(* IEC 61131-3 sources: plc-st-coding-agent/progress/evidence/f14_v14_remaining_20261113/jobs/codex_minimax-m27 (part 5) *)

(* ---- self-hard-03.raw_candidate_01.st ---- *)
(* ENGINEERING_CONTRACT
 * FIFO Queue with 8-slot compact array
 * [PUB001-PUB010] Core ops: popEn rising→remove first if count>0; pushEn rising→add pushItem if count<8
 *   Same-scan priority: pop executes BEFORE push; full→pop+push (net 0), empty→push-only (net +1)
 * [PUB011] Retention: count and fifo[1..8] state retained in VAR between scans
 * [PUB012] No AT located declarations
 * [PUB013-PUB015] Rising edge: each button triggers once per press; initial history=FALSE
 * [PUB016-PUB019] Same-scan semantics: full queue drains one slot then accepts push; empty queue accepts push only
 * [PUB020-PUB025] Array bounds: fifo[1..8], compact at end of scan: fifo[1..count] is logical queue FIFO order
 *   head=fifo[1] when non-empty, else 0; fifo[count+1..8] unspecified/unconstrained
 * [PUB026-PUB030] count∈[0,8], full↔count=8, empty↔count=0; success of push/pop updates count
 *)

(* CONTRACT_RULES [] *)

FUNCTION_BLOCK FB
VAR_INPUT
    pushEn    : BOOL;
    pushItem  : INT;
    popEn     : BOOL;
END_VAR
VAR_IN_OUT
    fifo      : ARRAY[1..8] OF INT;
END_VAR
VAR_OUTPUT
    count     : INT;
    full      : BOOL;
    empty     : BOOL;
    head      : INT;
END_VAR
VAR
    prev_pushEn : BOOL := FALSE;
    prev_popEn  : BOOL := FALSE;
    tmp_pushRising : BOOL;
    tmp_popRising  : BOOL;
    tmp_i       : INT;
END_VAR

    // Rising edge detection
    tmp_popRising  := popEn AND NOT prev_popEn;
    tmp_pushRising := pushEn AND NOT prev_pushEn;
    prev_popEn  := popEn;
    prev_pushEn := pushEn;

    // Execute in required order: pop first, then push
    // POP: non-empty queue only
    IF tmp_popRising AND count > 0 THEN
        FOR tmp_i := 1 TO count - 1 DO
            fifo[tmp_i] := fifo[tmp_i + 1];
        END_FOR;
        count := count - 1;
    END_IF;

    // PUSH: non-full queue only
    IF tmp_pushRising AND count < 8 THEN
        count := count + 1;
        fifo[count] := pushItem;
    END_IF;

    // Outputs
    full  := (count = 8);
    empty := (count = 0);
    IF empty THEN
        head := 0;
    ELSE
        head := fifo[1];
    END_IF;

END_FUNCTION_BLOCK

(* ---- self-hard-04.candidate_01.st ---- *)
(*
ENGINEERING_CONTRACT
==================
State retention & activation:
- leadPump: latches until demand=0 clears it; reset_input=demand<=0 PUB004
- lagPump: latches until demand<2 clears it; hold on same-scan no-rise PUB005
- runningCount: combinational, equals clipped demand every scan PUB001
Initialization:
- First positive demand after demand=0 selects shortest-run pump as leadPump (PUB010)
- First positive demand sets lagPump if demand>=2 (PUB011)
Rotation behavior:
- rotated=TRUE + main.runHours - MIN(runHours) > 50 → switch to shortest (PUB012)
- rotated=FALSE → never switch, even if hysteresis gap exists (PUB012)
- rotated is level-triggered, evaluated every scan with current main hours (PUB012)
Backup selection moments:
- Initial selection | leadPump change | runningCount increase → recompute lagPump (PUB026)
- Otherwise retain previous lagPump (PUB028)
Direction conflict: N/A (no opposite movements in this pump-selection task)
Units: runHours in LINT hours, 50-hour hysteresis threshold (PUB012)
*)
(* CONTRACT_RULES [] *)

FUNCTION_BLOCK FB
VAR_INPUT
    demand     : INT;
    runHours   : ARRAY[1..5] OF LINT;
    rotated    : BOOL;
END_VAR
VAR_OUTPUT
    leadPump   : INT := 0;
    lagPump    : INT := 0;
    runningCount : INT := 0;
END_VAR
VAR
    prevLeadPump    : INT := 0;
    prevLagPump     : INT := 0;
    prevRunningCount : INT := 0;
    prevClippedDemand : INT := 0;
    wasDemandZero   : BOOL := TRUE;
END_VAR

VAR
    clippedDemand : INT;
    tmp_i         : INT;
    tmp_minHours  : LINT;
    tmp_minPump   : INT;
    tmp_secondMinHours : LINT;
    tmp_secondMinPump  : INT;
    tmp_mainHoursDiff  : LINT;
END_VAR

    // PUB001: Clip demand to 0..5
    IF demand < 0 THEN
        clippedDemand := 0;
    ELSIF demand > 5 THEN
        clippedDemand := 5;
    ELSE
        clippedDemand := demand;
    END_IF;

    runningCount := clippedDemand;

    // Clear all outputs when demand <= 0
    IF clippedDemand = 0 THEN
        leadPump := 0;
        lagPump  := 0;
        prevLeadPump    := 0;
        prevLagPump     := 0;
        prevRunningCount := 0;
        prevClippedDemand := 0;
        wasDemandZero   := TRUE;
    ELSE
        // Find pump with minimum run hours (for hysteresis check and selection)
        tmp_minHours := runHours[1];
        tmp_minPump  := 1;
        FOR tmp_i := 2 TO 5 DO
            IF runHours[tmp_i] < tmp_minHours THEN
                tmp_minHours := runHours[tmp_i];
                tmp_minPump  := tmp_i;
            ELSIF runHours[tmp_i] = tmp_minHours AND tmp_i < tmp_minPump THEN
                tmp_minPump  := tmp_i;
            END_IF;
        END_FOR;

        // Determine if this is initial selection (first positive demand after zero)
        IF wasDemandZero THEN
            // Initial selection: pick shortest-run pump as main
            leadPump   := tmp_minPump;
            lagPump    := 0;
            wasDemandZero := FALSE;
        ELSE
            // Not initial selection: check for rotation request
            IF rotated AND prevLeadPump <> 0 THEN
                // Compute main pump's hours difference from minimum
                tmp_mainHoursDiff := runHours[prevLeadPump] - tmp_minHours;
                IF tmp_mainHoursDiff > 50 THEN
                    // Hysteresis satisfied: switch to shortest-run pump
                    leadPump := tmp_minPump;
                ELSE
                    // Keep current main pump
                    leadPump := prevLeadPump;
                END_IF;
            ELSE
                // No rotation request or no previous main: keep current main
                leadPump := prevLeadPump;
            END_IF;
        END_IF;

        // Backup pump selection (PUB026, PUB028)
        IF clippedDemand >= 2 THEN
            // Need backup pump
            // Recompute lagPump only on: initial, leadPump change, runningCount increase
            IF wasDemandZero OR leadPump <> prevLeadPump OR clippedDemand > prevClippedDemand THEN
                // Find second-minimum pump (excluding leadPump)
                tmp_secondMinHours := 16#7FFFFFFFFFFFFFFF; // Large LINT value
                tmp_secondMinPump  := 0;
                FOR tmp_i := 1 TO 5 DO
                    IF tmp_i = leadPump THEN
                        // Skip main pump
                    ELSE
                        IF runHours[tmp_i] < tmp_secondMinHours THEN
                            tmp_secondMinHours := runHours[tmp_i];
                            tmp_secondMinPump  := tmp_i;
                        ELSIF runHours[tmp_i] = tmp_secondMinHours AND tmp_i < tmp_secondMinPump THEN
                            tmp_secondMinPump  := tmp_i;
                        END_IF;
                    END_IF;
                END_FOR;
                lagPump := tmp_secondMinPump;
            ELSE
                // Retain previous backup pump
                lagPump := prevLagPump;
            END_IF;
        ELSE
            // Demand < 2: no backup pump
            lagPump := 0;
        END_IF;
    END_IF;

    // Update previous state for next scan
    prevLeadPump     := leadPump;
    prevLagPump      := lagPump;
    prevRunningCount := runningCount;
    prevClippedDemand := clippedDemand;

END_FUNCTION_BLOCK

(* ---- self-hard-04.candidate_03.st ---- *)
(*
ENGINEERING_CONTRACT
==================
State retention & activation:
- leadPump: latches until demand=0 clears it; reset_input=demand<=0 PUB004
- lagPump: latches until demand<2 clears it; hold on same-scan no-rise PUB005
- runningCount: combinational, equals clipped demand every scan PUB001
Initialization:
- First positive demand after demand=0 selects shortest-run pump as leadPump (PUB010)
- First positive demand sets lagPump if demand>=2 (PUB011)
Rotation behavior:
- rotated=TRUE + main.runHours - MIN(runHours) > 50 → switch to shortest (PUB012)
- rotated=FALSE → never switch, even if hysteresis gap exists (PUB012)
- rotated is level-triggered, evaluated every scan with current main hours (PUB012)
Backup selection moments:
- Initial selection | leadPump change | runningCount increase → recompute lagPump (PUB026)
- Otherwise retain previous lagPump (PUB028)
Direction conflict: N/A (no opposite movements in this pump-selection task)
Units: runHours in LINT hours, 50-hour hysteresis threshold (PUB012)
*)
(* CONTRACT_RULES [] *)

FUNCTION_BLOCK FB
VAR_INPUT
    demand     : INT;
    runHours   : ARRAY[1..5] OF LINT;
    rotated    : BOOL;
END_VAR
VAR_OUTPUT
    leadPump   : INT := 0;
    lagPump    : INT := 0;
    runningCount : INT := 0;
END_VAR
VAR
    prevLeadPump    : INT := 0;
    prevLagPump     : INT := 0;
    prevRunningCount : INT := 0;
    prevClippedDemand : INT := 0;
    wasDemandZero   : BOOL := TRUE;
    clippedDemand : INT;
    tmp_i         : INT;
    tmp_minHours  : LINT;
    tmp_minPump   : INT;
    tmp_secondMinHours : LINT;
    tmp_secondMinPump  : INT;
    tmp_mainHoursDiff  : LINT;
END_VAR

    // PUB001: Clip demand to 0..5
    IF demand < 0 THEN
        clippedDemand := 0;
    ELSIF demand > 5 THEN
        clippedDemand := 5;
    ELSE
        clippedDemand := demand;
    END_IF;

    runningCount := clippedDemand;

    // Clear all outputs when demand <= 0
    IF clippedDemand = 0 THEN
        leadPump := 0;
        lagPump  := 0;
        prevLeadPump    := 0;
        prevLagPump     := 0;
        prevRunningCount := 0;
        prevClippedDemand := 0;
        wasDemandZero   := TRUE;
    ELSE
        // Find pump with minimum run hours (for hysteresis check and selection)
        tmp_minHours := runHours[1];
        tmp_minPump  := 1;
        FOR tmp_i := 2 TO 5 DO
            IF runHours[tmp_i] < tmp_minHours THEN
                tmp_minHours := runHours[tmp_i];
                tmp_minPump  := tmp_i;
            ELSIF runHours[tmp_i] = tmp_minHours AND tmp_i < tmp_minPump THEN
                tmp_minPump  := tmp_i;
            END_IF;
        END_FOR;

        // Determine if this is initial selection (first positive demand after zero)
        IF wasDemandZero THEN
            // Initial selection: pick shortest-run pump as main
            leadPump   := tmp_minPump;
            lagPump    := 0;
            wasDemandZero := FALSE;
        ELSE
            // Not initial selection: check for rotation request
            IF rotated AND prevLeadPump <> 0 THEN
                // Compute main pump's hours difference from minimum
                tmp_mainHoursDiff := runHours[prevLeadPump] - tmp_minHours;
                IF tmp_mainHoursDiff > 50 THEN
                    // Hysteresis satisfied: switch to shortest-run pump
                    leadPump := tmp_minPump;
                ELSE
                    // Keep current main pump
                    leadPump := prevLeadPump;
                END_IF;
            ELSE
                // No rotation request or no previous main: keep current main
                leadPump := prevLeadPump;
            END_IF;
        END_IF;

        // Backup pump selection (PUB026, PUB028)
        IF clippedDemand >= 2 THEN
            // Need backup pump
            // Recompute lagPump only on: initial, leadPump change, runningCount increase
            IF wasDemandZero OR leadPump <> prevLeadPump OR clippedDemand > prevClippedDemand THEN
                // Find second-minimum pump (excluding leadPump)
                tmp_secondMinHours := 16#7FFFFFFFFFFFFFFF; // Large LINT value
                tmp_secondMinPump  := 0;
                FOR tmp_i := 1 TO 5 DO
                    IF tmp_i = leadPump THEN
                        // Skip main pump
                    ELSE
                        IF runHours[tmp_i] < tmp_secondMinHours THEN
                            tmp_secondMinHours := runHours[tmp_i];
                            tmp_secondMinPump  := tmp_i;
                        ELSIF runHours[tmp_i] = tmp_secondMinHours AND tmp_i < tmp_secondMinPump THEN
                            tmp_secondMinPump  := tmp_i;
                        END_IF;
                    END_IF;
                END_FOR;
                lagPump := tmp_secondMinPump;
            ELSE
                // Retain previous backup pump
                lagPump := prevLagPump;
            END_IF;
        ELSE
            // Demand < 2: no backup pump
            lagPump := 0;
        END_IF;
    END_IF;

    // Update previous state for next scan
    prevLeadPump     := leadPump;
    prevLagPump      := lagPump;
    prevRunningCount := runningCount;
    prevClippedDemand := clippedDemand;

END_FUNCTION_BLOCK

(* ---- self-hard-04.patch_base_02.st ---- *)
(*
ENGINEERING_CONTRACT
==================
State retention & activation:
- leadPump: latches until demand=0 clears it; reset_input=demand<=0 PUB004
- lagPump: latches until demand<2 clears it; hold on same-scan no-rise PUB005
- runningCount: combinational, equals clipped demand every scan PUB001
Initialization:
- First positive demand after demand=0 selects shortest-run pump as leadPump (PUB010)
- First positive demand sets lagPump if demand>=2 (PUB011)
Rotation behavior:
- rotated=TRUE + main.runHours - MIN(runHours) > 50 → switch to shortest (PUB012)
- rotated=FALSE → never switch, even if hysteresis gap exists (PUB012)
- rotated is level-triggered, evaluated every scan with current main hours (PUB012)
Backup selection moments:
- Initial selection | leadPump change | runningCount increase → recompute lagPump (PUB026)
- Otherwise retain previous lagPump (PUB028)
Direction conflict: N/A (no opposite movements in this pump-selection task)
Units: runHours in LINT hours, 50-hour hysteresis threshold (PUB012)
*)
(* CONTRACT_RULES [] *)

FUNCTION_BLOCK FB
VAR_INPUT
    demand     : INT;
    runHours   : ARRAY[1..5] OF LINT;
    rotated    : BOOL;
END_VAR
VAR_OUTPUT
    leadPump   : INT := 0;
    lagPump    : INT := 0;
    runningCount : INT := 0;
END_VAR
VAR
    prevLeadPump    : INT := 0;
    prevLagPump     : INT := 0;
    prevRunningCount : INT := 0;
    prevClippedDemand : INT := 0;
    wasDemandZero   : BOOL := TRUE;
END_VAR

VAR
    clippedDemand : INT;
    tmp_i         : INT;
    tmp_minHours  : LINT;
    tmp_minPump   : INT;
    tmp_secondMinHours : LINT;
    tmp_secondMinPump  : INT;
    tmp_mainHoursDiff  : LINT;
END_VAR

    // PUB001: Clip demand to 0..5
    IF demand < 0 THEN
        clippedDemand := 0;
    ELSIF demand > 5 THEN
        clippedDemand := 5;
    ELSE
        clippedDemand := demand;
    END_IF;

    runningCount := clippedDemand;

    // Clear all outputs when demand <= 0
    IF clippedDemand = 0 THEN
        leadPump := 0;
        lagPump  := 0;
        prevLeadPump    := 0;
        prevLagPump     := 0;
        prevRunningCount := 0;
        prevClippedDemand := 0;
        wasDemandZero   := TRUE;
    ELSE
        // Find pump with minimum run hours (for hysteresis check and selection)
        tmp_minHours := runHours[1];
        tmp_minPump  := 1;
        FOR tmp_i := 2 TO 5 DO
            IF runHours[tmp_i] < tmp_minHours THEN
                tmp_minHours := runHours[tmp_i];
                tmp_minPump  := tmp_i;
            ELSIF runHours[tmp_i] = tmp_minHours AND tmp_i < tmp_minPump THEN
                tmp_minPump  := tmp_i;
            END_IF;
        END_FOR;

        // Determine if this is initial selection (first positive demand after zero)
        IF wasDemandZero THEN
            // Initial selection: pick shortest-run pump as main
            leadPump   := tmp_minPump;
            lagPump    := 0;
            wasDemandZero := FALSE;
        ELSE
            // Not initial selection: check for rotation request
            IF rotated AND prevLeadPump <> 0 THEN
                // Compute main pump's hours difference from minimum
                tmp_mainHoursDiff := runHours[prevLeadPump] - tmp_minHours;
                IF tmp_mainHoursDiff > 50 THEN
                    // Hysteresis satisfied: switch to shortest-run pump
                    leadPump := tmp_minPump;
                ELSE
                    // Keep current main pump
                    leadPump := prevLeadPump;
                END_IF;
            ELSE
                // No rotation request or no previous main: keep current main
                leadPump := prevLeadPump;
            END_IF;
        END_IF;

        // Backup pump selection (PUB026, PUB028)
        IF clippedDemand >= 2 THEN
            // Need backup pump
            // Recompute lagPump only on: initial, leadPump change, runningCount increase
            IF wasDemandZero OR leadPump <> prevLeadPump OR clippedDemand > prevClippedDemand THEN
                // Find second-minimum pump (excluding leadPump)
                tmp_secondMinHours := 16#7FFFFFFFFFFFFFFF; // Large LINT value
                tmp_secondMinPump  := 0;
                FOR tmp_i := 1 TO 5 DO
                    IF tmp_i = leadPump THEN
                        // Skip main pump
                    ELSE
                        IF runHours[tmp_i] < tmp_secondMinHours THEN
                            tmp_secondMinHours := runHours[tmp_i];
                            tmp_secondMinPump  := tmp_i;
                        ELSIF runHours[tmp_i] = tmp_secondMinHours AND tmp_i < tmp_secondMinPump THEN
                            tmp_secondMinPump  := tmp_i;
                        END_IF;
                    END_IF;
                END_FOR;
                lagPump := tmp_secondMinPump;
            ELSE
                // Retain previous backup pump
                lagPump := prevLagPump;
            END_IF;
        ELSE
            // Demand < 2: no backup pump
            lagPump := 0;
        END_IF;
    END_IF;

    // Update previous state for next scan
    prevLeadPump     := leadPump;
    prevLagPump      := lagPump;
    prevRunningCount := runningCount;
    prevClippedDemand := clippedDemand;

END_FUNCTION_BLOCK

(* ---- self-hard-04.patch_base_03.st ---- *)
(*
ENGINEERING_CONTRACT
==================
State retention & activation:
- leadPump: latches until demand=0 clears it; reset_input=demand<=0 PUB004
- lagPump: latches until demand<2 clears it; hold on same-scan no-rise PUB005
- runningCount: combinational, equals clipped demand every scan PUB001
Initialization:
- First positive demand after demand=0 selects shortest-run pump as leadPump (PUB010)
- First positive demand sets lagPump if demand>=2 (PUB011)
Rotation behavior:
- rotated=TRUE + main.runHours - MIN(runHours) > 50 → switch to shortest (PUB012)
- rotated=FALSE → never switch, even if hysteresis gap exists (PUB012)
- rotated is level-triggered, evaluated every scan with current main hours (PUB012)
Backup selection moments:
- Initial selection | leadPump change | runningCount increase → recompute lagPump (PUB026)
- Otherwise retain previous lagPump (PUB028)
Direction conflict: N/A (no opposite movements in this pump-selection task)
Units: runHours in LINT hours, 50-hour hysteresis threshold (PUB012)
*)
(* CONTRACT_RULES [] *)

FUNCTION_BLOCK FB
VAR_INPUT
    demand     : INT;
    runHours   : ARRAY[1..5] OF LINT;
    rotated    : BOOL;
END_VAR
VAR_OUTPUT
    leadPump   : INT := 0;
    lagPump    : INT := 0;
    runningCount : INT := 0;
END_VAR
VAR
    prevLeadPump    : INT := 0;
    prevLagPump     : INT := 0;
    prevRunningCount : INT := 0;
    prevClippedDemand : INT := 0;
    wasDemandZero   : BOOL := TRUE;
END_VAR

VAR
    clippedDemand : INT;
    tmp_i         : INT;
    tmp_minHours  : LINT;
    tmp_minPump   : INT;
    tmp_secondMinHours : LINT;
    tmp_secondMinPump  : INT;
    tmp_mainHoursDiff  : LINT;
END_VAR

    // PUB001: Clip demand to 0..5
    IF demand < 0 THEN
        clippedDemand := 0;
    ELSIF demand > 5 THEN
        clippedDemand := 5;
    ELSE
        clippedDemand := demand;
    END_IF;

    runningCount := clippedDemand;

    // Clear all outputs when demand <= 0
    IF clippedDemand = 0 THEN
        leadPump := 0;
        lagPump  := 0;
        prevLeadPump    := 0;
        prevLagPump     := 0;
        prevRunningCount := 0;
        prevClippedDemand := 0;
        wasDemandZero   := TRUE;
    ELSE
        // Find pump with minimum run hours (for hysteresis check and selection)
        tmp_minHours := runHours[1];
        tmp_minPump  := 1;
        FOR tmp_i := 2 TO 5 DO
            IF runHours[tmp_i] < tmp_minHours THEN
                tmp_minHours := runHours[tmp_i];
                tmp_minPump  := tmp_i;
            ELSIF runHours[tmp_i] = tmp_minHours AND tmp_i < tmp_minPump THEN
                tmp_minPump  := tmp_i;
            END_IF;
        END_FOR;

        // Determine if this is initial selection (first positive demand after zero)
        IF wasDemandZero THEN
            // Initial selection: pick shortest-run pump as main
            leadPump   := tmp_minPump;
            lagPump    := 0;
            wasDemandZero := FALSE;
        ELSE
            // Not initial selection: check for rotation request
            IF rotated AND prevLeadPump <> 0 THEN
                // Compute main pump's hours difference from minimum
                tmp_mainHoursDiff := runHours[prevLeadPump] - tmp_minHours;
                IF tmp_mainHoursDiff > 50 THEN
                    // Hysteresis satisfied: switch to shortest-run pump
                    leadPump := tmp_minPump;
                ELSE
                    // Keep current main pump
                    leadPump := prevLeadPump;
                END_IF;
            ELSE
                // No rotation request or no previous main: keep current main
                leadPump := prevLeadPump;
            END_IF;
        END_IF;

        // Backup pump selection (PUB026, PUB028)
        IF clippedDemand >= 2 THEN
            // Need backup pump
            // Recompute lagPump only on: initial, leadPump change, runningCount increase
            IF wasDemandZero OR leadPump <> prevLeadPump OR clippedDemand > prevClippedDemand THEN
                // Find second-minimum pump (excluding leadPump)
                tmp_secondMinHours := 16#7FFFFFFFFFFFFFFF; // Large LINT value
                tmp_secondMinPump  := 0;
                FOR tmp_i := 1 TO 5 DO
                    IF tmp_i = leadPump THEN
                        // Skip main pump
                    ELSE
                        IF runHours[tmp_i] < tmp_secondMinHours THEN
                            tmp_secondMinHours := runHours[tmp_i];
                            tmp_secondMinPump  := tmp_i;
                        ELSIF runHours[tmp_i] = tmp_secondMinHours AND tmp_i < tmp_secondMinPump THEN
                            tmp_secondMinPump  := tmp_i;
                        END_IF;
                    END_IF;
                END_FOR;
                lagPump := tmp_secondMinPump;
            ELSE
                // Retain previous backup pump
                lagPump := prevLagPump;
            END_IF;
        ELSE
            // Demand < 2: no backup pump
            lagPump := 0;
        END_IF;
    END_IF;

    // Update previous state for next scan
    prevLeadPump     := leadPump;
    prevLagPump      := lagPump;
    prevRunningCount := runningCount;
    prevClippedDemand := clippedDemand;

END_FUNCTION_BLOCK

(* ---- self-hard-04.patch_base_04.st ---- *)
(*
ENGINEERING_CONTRACT
==================
State retention & activation:
- leadPump: latches until demand=0 clears it; reset_input=demand<=0 PUB004
- lagPump: latches until demand<2 clears it; hold on same-scan no-rise PUB005
- runningCount: combinational, equals clipped demand every scan PUB001
Initialization:
- First positive demand after demand=0 selects shortest-run pump as leadPump (PUB010)
- First positive demand sets lagPump if demand>=2 (PUB011)
Rotation behavior:
- rotated=TRUE + main.runHours - MIN(runHours) > 50 → switch to shortest (PUB012)
- rotated=FALSE → never switch, even if hysteresis gap exists (PUB012)
- rotated is level-triggered, evaluated every scan with current main hours (PUB012)
Backup selection moments:
- Initial selection | leadPump change | runningCount increase → recompute lagPump (PUB026)
- Otherwise retain previous lagPump (PUB028)
Direction conflict: N/A (no opposite movements in this pump-selection task)
Units: runHours in LINT hours, 50-hour hysteresis threshold (PUB012)
*)
(* CONTRACT_RULES [] *)

FUNCTION_BLOCK FB
VAR_INPUT
    demand     : INT;
    runHours   : ARRAY[1..5] OF LINT;
    rotated    : BOOL;
END_VAR
VAR_OUTPUT
    leadPump   : INT := 0;
    lagPump    : INT := 0;
    runningCount : INT := 0;
END_VAR
VAR
    prevLeadPump    : INT := 0;
    prevLagPump     : INT := 0;
    prevRunningCount : INT := 0;
    prevClippedDemand : INT := 0;
    wasDemandZero   : BOOL := TRUE;
    clippedDemand : INT;
    tmp_i         : INT;
    tmp_minHours  : LINT;
    tmp_minPump   : INT;
    tmp_secondMinHours : LINT;
    tmp_secondMinPump  : INT;
    tmp_mainHoursDiff  : LINT;
END_VAR

    // PUB001: Clip demand to 0..5
    IF demand < 0 THEN
        clippedDemand := 0;
    ELSIF demand > 5 THEN
        clippedDemand := 5;
    ELSE
        clippedDemand := demand;
    END_IF;

    runningCount := clippedDemand;

    // Clear all outputs when demand <= 0
    IF clippedDemand = 0 THEN
        leadPump := 0;
        lagPump  := 0;
        prevLeadPump    := 0;
        prevLagPump     := 0;
        prevRunningCount := 0;
        prevClippedDemand := 0;
        wasDemandZero   := TRUE;
    ELSE
        // Find pump with minimum run hours (for hysteresis check and selection)
        tmp_minHours := runHours[1];
        tmp_minPump  := 1;
        FOR tmp_i := 2 TO 5 DO
            IF runHours[tmp_i] < tmp_minHours THEN
                tmp_minHours := runHours[tmp_i];
                tmp_minPump  := tmp_i;
            ELSIF runHours[tmp_i] = tmp_minHours AND tmp_i < tmp_minPump THEN
                tmp_minPump  := tmp_i;
            END_IF;
        END_FOR;

        // Determine if this is initial selection (first positive demand after zero)
        IF wasDemandZero THEN
            // Initial selection: pick shortest-run pump as main
            leadPump   := tmp_minPump;
            lagPump    := 0;
            wasDemandZero := FALSE;
        ELSE
            // Not initial selection: check for rotation request
            IF rotated AND prevLeadPump <> 0 THEN
                // Compute main pump's hours difference from minimum
                tmp_mainHoursDiff := runHours[prevLeadPump] - tmp_minHours;
                IF tmp_mainHoursDiff > 50 THEN
                    // Hysteresis satisfied: switch to shortest-run pump
                    leadPump := tmp_minPump;
                ELSE
                    // Keep current main pump
                    leadPump := prevLeadPump;
                END_IF;
            ELSE
                // No rotation request or no previous main: keep current main
                leadPump := prevLeadPump;
            END_IF;
        END_IF;

        // Backup pump selection (PUB026, PUB028)
        IF clippedDemand >= 2 THEN
            // Need backup pump
            // Recompute lagPump only on: initial, leadPump change, runningCount increase
            IF wasDemandZero OR leadPump <> prevLeadPump OR clippedDemand > prevClippedDemand THEN
                // Find second-minimum pump (excluding leadPump)
                tmp_secondMinHours := 16#7FFFFFFFFFFFFFFF; // Large LINT value
                tmp_secondMinPump  := 0;
                FOR tmp_i := 1 TO 5 DO
                    IF tmp_i = leadPump THEN
                        // Skip main pump
                    ELSE
                        IF runHours[tmp_i] < tmp_secondMinHours THEN
                            tmp_secondMinHours := runHours[tmp_i];
                            tmp_secondMinPump  := tmp_i;
                        ELSIF runHours[tmp_i] = tmp_secondMinHours AND tmp_i < tmp_secondMinPump THEN
                            tmp_secondMinPump  := tmp_i;
                        END_IF;
                    END_IF;
                END_FOR;
                lagPump := tmp_secondMinPump;
            ELSE
                // Retain previous backup pump
                lagPump := prevLagPump;
            END_IF;
        ELSE
            // Demand < 2: no backup pump
            lagPump := 0;
        END_IF;
    END_IF;

    // Update previous state for next scan
    prevLeadPump     := leadPump;
    prevLagPump      := lagPump;
    prevRunningCount := runningCount;
    prevClippedDemand := clippedDemand;

END_FUNCTION_BLOCK

(* ---- self-hard-04.raw_candidate_01.st ---- *)
(*
ENGINEERING_CONTRACT
==================
State retention & activation:
- leadPump: latches until demand=0 clears it; reset_input=demand<=0 PUB004
- lagPump: latches until demand<2 clears it; hold on same-scan no-rise PUB005
- runningCount: combinational, equals clipped demand every scan PUB001
Initialization:
- First positive demand after demand=0 selects shortest-run pump as leadPump (PUB010)
- First positive demand sets lagPump if demand>=2 (PUB011)
Rotation behavior:
- rotated=TRUE + main.runHours - MIN(runHours) > 50 → switch to shortest (PUB012)
- rotated=FALSE → never switch, even if hysteresis gap exists (PUB012)
- rotated is level-triggered, evaluated every scan with current main hours (PUB012)
Backup selection moments:
- Initial selection | leadPump change | runningCount increase → recompute lagPump (PUB026)
- Otherwise retain previous lagPump (PUB028)
Direction conflict: N/A (no opposite movements in this pump-selection task)
Units: runHours in LINT hours, 50-hour hysteresis threshold (PUB012)
*)
(* CONTRACT_RULES [] *)

FUNCTION_BLOCK FB
VAR_INPUT
    demand     : INT;
    runHours   : ARRAY[1..5] OF LINT;
    rotated    : BOOL;
END_VAR
VAR_OUTPUT
    leadPump   : INT := 0;
    lagPump    : INT := 0;
    runningCount : INT := 0;
END_VAR
VAR
    prevLeadPump    : INT := 0;
    prevLagPump     : INT := 0;
    prevRunningCount : INT := 0;
    prevClippedDemand : INT := 0;
    wasDemandZero   : BOOL := TRUE;
END_VAR

VAR
    clippedDemand : INT;
    tmp_i         : INT;
    tmp_minHours  : LINT;
    tmp_minPump   : INT;
    tmp_secondMinHours : LINT;
    tmp_secondMinPump  : INT;
    tmp_mainHoursDiff  : LINT;
END_VAR

    // PUB001: Clip demand to 0..5
    IF demand < 0 THEN
        clippedDemand := 0;
    ELSIF demand > 5 THEN
        clippedDemand := 5;
    ELSE
        clippedDemand := demand;
    END_IF;

    runningCount := clippedDemand;

    // Clear all outputs when demand <= 0
    IF clippedDemand = 0 THEN
        leadPump := 0;
        lagPump  := 0;
        prevLeadPump    := 0;
        prevLagPump     := 0;
        prevRunningCount := 0;
        prevClippedDemand := 0;
        wasDemandZero   := TRUE;
    ELSE
        // Find pump with minimum run hours (for hysteresis check and selection)
        tmp_minHours := runHours[1];
        tmp_minPump  := 1;
        FOR tmp_i := 2 TO 5 DO
            IF runHours[tmp_i] < tmp_minHours THEN
                tmp_minHours := runHours[tmp_i];
                tmp_minPump  := tmp_i;
            ELSIF runHours[tmp_i] = tmp_minHours AND tmp_i < tmp_minPump THEN
                tmp_minPump  := tmp_i;
            END_IF;
        END_FOR;

        // Determine if this is initial selection (first positive demand after zero)
        IF wasDemandZero THEN
            // Initial selection: pick shortest-run pump as main
            leadPump   := tmp_minPump;
            lagPump    := 0;
            wasDemandZero := FALSE;
        ELSE
            // Not initial selection: check for rotation request
            IF rotated AND prevLeadPump <> 0 THEN
                // Compute main pump's hours difference from minimum
                tmp_mainHoursDiff := runHours[prevLeadPump] - tmp_minHours;
                IF tmp_mainHoursDiff > 50 THEN
                    // Hysteresis satisfied: switch to shortest-run pump
                    leadPump := tmp_minPump;
                ELSE
                    // Keep current main pump
                    leadPump := prevLeadPump;
                END_IF;
            ELSE
                // No rotation request or no previous main: keep current main
                leadPump := prevLeadPump;
            END_IF;
        END_IF;

        // Backup pump selection (PUB026, PUB028)
        IF clippedDemand >= 2 THEN
            // Need backup pump
            // Recompute lagPump only on: initial, leadPump change, runningCount increase
            IF wasDemandZero OR leadPump <> prevLeadPump OR clippedDemand > prevClippedDemand THEN
                // Find second-minimum pump (excluding leadPump)
                tmp_secondMinHours := 16#7FFFFFFFFFFFFFFF; // Large LINT value
                tmp_secondMinPump  := 0;
                FOR tmp_i := 1 TO 5 DO
                    IF tmp_i = leadPump THEN
                        // Skip main pump
                    ELSE
                        IF runHours[tmp_i] < tmp_secondMinHours THEN
                            tmp_secondMinHours := runHours[tmp_i];
                            tmp_secondMinPump  := tmp_i;
                        ELSIF runHours[tmp_i] = tmp_secondMinHours AND tmp_i < tmp_secondMinPump THEN
                            tmp_secondMinPump  := tmp_i;
                        END_IF;
                    END_IF;
                END_FOR;
                lagPump := tmp_secondMinPump;
            ELSE
                // Retain previous backup pump
                lagPump := prevLagPump;
            END_IF;
        ELSE
            // Demand < 2: no backup pump
            lagPump := 0;
        END_IF;
    END_IF;

    // Update previous state for next scan
    prevLeadPump     := leadPump;
    prevLagPump      := lagPump;
    prevRunningCount := runningCount;
    prevClippedDemand := clippedDemand;

END_FUNCTION_BLOCK

(* ---- self-hard-04.raw_candidate_03.st ---- *)
(*
ENGINEERING_CONTRACT
==================
State retention & activation:
- leadPump: latches until demand=0 clears it; reset_input=demand<=0 PUB004
- lagPump: latches until demand<2 clears it; hold on same-scan no-rise PUB005
- runningCount: combinational, equals clipped demand every scan PUB001
Initialization:
- First positive demand after demand=0 selects shortest-run pump as leadPump (PUB010)
- First positive demand sets lagPump if demand>=2 (PUB011)
Rotation behavior:
- rotated=TRUE + main.runHours - MIN(runHours) > 50 → switch to shortest (PUB012)
- rotated=FALSE → never switch, even if hysteresis gap exists (PUB012)
- rotated is level-triggered, evaluated every scan with current main hours (PUB012)
Backup selection moments:
- Initial selection | leadPump change | runningCount increase → recompute lagPump (PUB026)
- Otherwise retain previous lagPump (PUB028)
Direction conflict: N/A (no opposite movements in this pump-selection task)
Units: runHours in LINT hours, 50-hour hysteresis threshold (PUB012)
*)
(* CONTRACT_RULES [] *)

FUNCTION_BLOCK FB
VAR_INPUT
    demand     : INT;
    runHours   : ARRAY[1..5] OF LINT;
    rotated    : BOOL;
END_VAR
VAR_OUTPUT
    leadPump   : INT := 0;
    lagPump    : INT := 0;
    runningCount : INT := 0;
END_VAR
VAR
    prevLeadPump    : INT := 0;
    prevLagPump     : INT := 0;
    prevRunningCount : INT := 0;
    prevClippedDemand : INT := 0;
    wasDemandZero   : BOOL := TRUE;
    clippedDemand : INT;
    tmp_i         : INT;
    tmp_minHours  : LINT;
    tmp_minPump   : INT;
    tmp_secondMinHours : LINT;
    tmp_secondMinPump  : INT;
    tmp_mainHoursDiff  : LINT;
END_VAR

    // PUB001: Clip demand to 0..5
    IF demand < 0 THEN
        clippedDemand := 0;
    ELSIF demand > 5 THEN
        clippedDemand := 5;
    ELSE
        clippedDemand := demand;
    END_IF;

    runningCount := clippedDemand;

    // Clear all outputs when demand <= 0
    IF clippedDemand = 0 THEN
        leadPump := 0;
        lagPump  := 0;
        prevLeadPump    := 0;
        prevLagPump     := 0;
        prevRunningCount := 0;
        prevClippedDemand := 0;
        wasDemandZero   := TRUE;
    ELSE
        // Find pump with minimum run hours (for hysteresis check and selection)
        tmp_minHours := runHours[1];
        tmp_minPump  := 1;
        FOR tmp_i := 2 TO 5 DO
            IF runHours[tmp_i] < tmp_minHours THEN
                tmp_minHours := runHours[tmp_i];
                tmp_minPump  := tmp_i;
            ELSIF runHours[tmp_i] = tmp_minHours AND tmp_i < tmp_minPump THEN
                tmp_minPump  := tmp_i;
            END_IF;
        END_FOR;

        // Determine if this is initial selection (first positive demand after zero)
        IF wasDemandZero THEN
            // Initial selection: pick shortest-run pump as main
            leadPump   := tmp_minPump;
            lagPump    := 0;
            wasDemandZero := FALSE;
        ELSE
            // Not initial selection: check for rotation request
            IF rotated AND prevLeadPump <> 0 THEN
                // Compute main pump's hours difference from minimum
                tmp_mainHoursDiff := runHours[prevLeadPump] - tmp_minHours;
                IF tmp_mainHoursDiff > 50 THEN
                    // Hysteresis satisfied: switch to shortest-run pump
                    leadPump := tmp_minPump;
                ELSE
                    // Keep current main pump
                    leadPump := prevLeadPump;
                END_IF;
            ELSE
                // No rotation request or no previous main: keep current main
                leadPump := prevLeadPump;
            END_IF;
        END_IF;

        // Backup pump selection (PUB026, PUB028)
        IF clippedDemand >= 2 THEN
            // Need backup pump
            // Recompute lagPump only on: initial, leadPump change, runningCount increase
            IF wasDemandZero OR leadPump <> prevLeadPump OR clippedDemand > prevClippedDemand THEN
                // Find second-minimum pump (excluding leadPump)
                tmp_secondMinHours := 16#7FFFFFFFFFFFFFFF; // Large LINT value
                tmp_secondMinPump  := 0;
                FOR tmp_i := 1 TO 5 DO
                    IF tmp_i = leadPump THEN
                        // Skip main pump
                    ELSE
                        IF runHours[tmp_i] < tmp_secondMinHours THEN
                            tmp_secondMinHours := runHours[tmp_i];
                            tmp_secondMinPump  := tmp_i;
                        ELSIF runHours[tmp_i] = tmp_secondMinHours AND tmp_i < tmp_secondMinPump THEN
                            tmp_secondMinPump  := tmp_i;
                        END_IF;
                    END_IF;
                END_FOR;
                lagPump := tmp_secondMinPump;
            ELSE
                // Retain previous backup pump
                lagPump := prevLagPump;
            END_IF;
        ELSE
            // Demand < 2: no backup pump
            lagPump := 0;
        END_IF;
    END_IF;

    // Update previous state for next scan
    prevLeadPump     := leadPump;
    prevLagPump      := lagPump;
    prevRunningCount := runningCount;
    prevClippedDemand := clippedDemand;

END_FUNCTION_BLOCK

(* ---- self-hard-05.candidate_01.st ---- *)
FUNCTION_BLOCK FB
VAR_INPUT
    runRequest  : BOOL;
    flameOK     : BOOL;
    o2Valid     : BOOL;
    o2PV        : REAL;
    baseAir     : REAL;
    resetBtn    : BOOL;
END_VAR
VAR_OUTPUT
    fuelPermit  : BOOL;
    trimEnable  : BOOL;
    airTrim     : REAL;
    airCommand  : REAL;
    tripLatched : BOOL;
    o2Fault     : BOOL;
END_VAR
VAR
    tmp_reset_rising : BOOL;
    tmp_trip_set     : BOOL;
END_VAR
(* ENGINEERING_CONTRACT
 * Output: tripLatched
 *   - SET:   runRequest=TRUE AND flameOK=FALSE  → same scan, no delay  [PUB001]
 *   - HOLD:  once set, retained across scans until valid reset edge     [PUB016]
 *   - RESET: rising(resetBtn) AND runRequest=FALSE AND flameOK=FALSE    [PUB016]
 *   - Edge-only reset; hold/rescan does NOT clear; press without edge does NOT clear
 * Output: fuelPermit
 *   - Activation:   runRequest AND flameOK AND NOT tripLatched          [PUB003]
 *   - Retention:    none — combinational, 0 when tripLatched           [PUB003]
 *   - Deactivation: tripLatched rising sets to FALSE; also 0 when any input low [PUB003]
 *   - Units: BOOLEAN
 * Output: trimEnable
 *   - Activation:   fuelPermit=TRUE AND o2Fault=FALSE                    [PUB008]
 *   - Retention:    none — combinational, 0 when o2Fault                [PUB008]
 *   - Deactivation: o2Fault rising (invalid/range)                      [PUB008]
 * Output: airTrim
 *   - Activation:   trimEnable with formula 2.0*(2.0-o2PV), clamp ±10   [PUB005]
 *   - Retention:    0.0 when trimEnable=FALSE (no residual)             [PUB010]
 *   - Units: % offset, clamped [-10,+10]
 * Output: airCommand
 *   - Activation:   baseAir+airTrim clamped [0,100] when fuelPermit=TRUE [PUB006]
 *   - Retention:    0.0 when fuelPermit=FALSE                           [PUB005]
 *   - Units: % absolute, clamped [0,100]; baseAir may be outside range [PUB006]
 * Output: o2Fault
 *   - Activation:   NOT o2Valid OR o2PV<0 OR o2PV>21                    [PUB009]
 *   - Retention:    combinational; does not inhibit fuelPermit          [PUB009]
 * Same-scan priority: trip set, fuelPermit, trimEnable/o2Fault, airTrim, airCommand
 * CONTRACT_RULES []
 *)
    // Detect rising edge of reset button (edge-only reset per PUB016)
    tmp_reset_rising := resetBtn AND NOT tmp_reset_rising;

    // Trip latch: set when running without flame, hold until valid reset edge
    tmp_trip_set := runRequest AND NOT flameOK;
    IF tmp_trip_set THEN
        tripLatched := TRUE;
    ELSIF tmp_reset_rising AND NOT runRequest AND NOT flameOK THEN
        tripLatched := FALSE;
    END_IF;

    // Fuel permit: requires run, flame, and no trip
    fuelPermit := runRequest AND flameOK AND NOT tripLatched;

    // O2 fault detection
    o2Fault := NOT o2Valid OR o2PV < 0.0 OR o2PV > 21.0;

    // Trim enable: fuel permit without O2 fault
    trimEnable := fuelPermit AND NOT o2Fault;

    // Air trim: 2.0*(2.0-o2PV), clamped to [-10, +10]; forced 0 when disabled
    IF trimEnable THEN
        airTrim := 2.0 * (2.0 - o2PV);
        IF airTrim > 10.0 THEN
            airTrim := 10.0;
        ELSIF airTrim < -10.0 THEN
            airTrim := -10.0;
        END_IF;
    ELSE
        airTrim := 0.0;
    END_IF;

    // Air command: base + trim, clamped [0,100]; forced 0 when no fuel permit
    IF fuelPermit THEN
        airCommand := baseAir + airTrim;
        IF airCommand > 100.0 THEN
            airCommand := 100.0;
        ELSIF airCommand < 0.0 THEN
            airCommand := 0.0;
        END_IF;
    ELSE
        airCommand := 0.0;
    END_IF;
END_FUNCTION_BLOCK

(* ---- self-hard-05.patch_base_02.st ---- *)
FUNCTION_BLOCK FB
VAR_INPUT
    runRequest  : BOOL;
    flameOK     : BOOL;
    o2Valid     : BOOL;
    o2PV        : REAL;
    baseAir     : REAL;
    resetBtn    : BOOL;
END_VAR
VAR_OUTPUT
    fuelPermit  : BOOL;
    trimEnable  : BOOL;
    airTrim     : REAL;
    airCommand  : REAL;
    tripLatched : BOOL;
    o2Fault     : BOOL;
END_VAR
VAR
    tmp_reset_rising : BOOL;
    tmp_trip_set     : BOOL;
END_VAR
(* ENGINEERING_CONTRACT
 * Output: tripLatched
 *   - SET:   runRequest=TRUE AND flameOK=FALSE  → same scan, no delay  [PUB001]
 *   - HOLD:  once set, retained across scans until valid reset edge     [PUB016]
 *   - RESET: rising(resetBtn) AND runRequest=FALSE AND flameOK=FALSE    [PUB016]
 *   - Edge-only reset; hold/rescan does NOT clear; press without edge does NOT clear
 * Output: fuelPermit
 *   - Activation:   runRequest AND flameOK AND NOT tripLatched          [PUB003]
 *   - Retention:    none — combinational, 0 when tripLatched           [PUB003]
 *   - Deactivation: tripLatched rising sets to FALSE; also 0 when any input low [PUB003]
 *   - Units: BOOLEAN
 * Output: trimEnable
 *   - Activation:   fuelPermit=TRUE AND o2Fault=FALSE                    [PUB008]
 *   - Retention:    none — combinational, 0 when o2Fault                [PUB008]
 *   - Deactivation: o2Fault rising (invalid/range)                      [PUB008]
 * Output: airTrim
 *   - Activation:   trimEnable with formula 2.0*(2.0-o2PV), clamp ±10   [PUB005]
 *   - Retention:    0.0 when trimEnable=FALSE (no residual)             [PUB010]
 *   - Units: % offset, clamped [-10,+10]
 * Output: airCommand
 *   - Activation:   baseAir+airTrim clamped [0,100] when fuelPermit=TRUE [PUB006]
 *   - Retention:    0.0 when fuelPermit=FALSE                           [PUB005]
 *   - Units: % absolute, clamped [0,100]; baseAir may be outside range [PUB006]
 * Output: o2Fault
 *   - Activation:   NOT o2Valid OR o2PV<0 OR o2PV>21                    [PUB009]
 *   - Retention:    combinational; does not inhibit fuelPermit          [PUB009]
 * Same-scan priority: trip set, fuelPermit, trimEnable/o2Fault, airTrim, airCommand
 * CONTRACT_RULES []
 *)
    // Detect rising edge of reset button (edge-only reset per PUB016)
    tmp_reset_rising := resetBtn AND NOT tmp_reset_rising;

    // Trip latch: set when running without flame, hold until valid reset edge
    tmp_trip_set := runRequest AND NOT flameOK;
    IF tmp_trip_set THEN
        tripLatched := TRUE;
    ELSIF tmp_reset_rising AND NOT runRequest AND NOT flameOK THEN
        tripLatched := FALSE;
    END_IF;

    // Fuel permit: requires run, flame, and no trip
    fuelPermit := runRequest AND flameOK AND NOT tripLatched;

    // O2 fault detection
    o2Fault := NOT o2Valid OR o2PV < 0.0 OR o2PV > 21.0;

    // Trim enable: fuel permit without O2 fault
    trimEnable := fuelPermit AND NOT o2Fault;

    // Air trim: 2.0*(2.0-o2PV), clamped to [-10, +10]; forced 0 when disabled
    IF trimEnable THEN
        airTrim := 2.0 * (2.0 - o2PV);
        IF airTrim > 10.0 THEN
            airTrim := 10.0;
        ELSIF airTrim < -10.0 THEN
            airTrim := -10.0;
        END_IF;
    ELSE
        airTrim := 0.0;
    END_IF;

    // Air command: base + trim, clamped [0,100]; forced 0 when no fuel permit
    IF fuelPermit THEN
        airCommand := baseAir + airTrim;
        IF airCommand > 100.0 THEN
            airCommand := 100.0;
        ELSIF airCommand < 0.0 THEN
            airCommand := 0.0;
        END_IF;
    ELSE
        airCommand := 0.0;
    END_IF;
END_FUNCTION_BLOCK

(* ---- self-hard-05.patch_base_03.st ---- *)
FUNCTION_BLOCK FB
VAR_INPUT
    runRequest  : BOOL;
    flameOK     : BOOL;
    o2Valid     : BOOL;
    o2PV        : REAL;
    baseAir     : REAL;
    resetBtn    : BOOL;
END_VAR
VAR_OUTPUT
    fuelPermit  : BOOL;
    trimEnable  : BOOL;
    airTrim     : REAL;
    airCommand  : REAL;
    tripLatched : BOOL;
    o2Fault     : BOOL;
END_VAR
VAR
    tmp_reset_rising : BOOL;
    tmp_trip_set     : BOOL;
END_VAR
(* ENGINEERING_CONTRACT
 * Output: tripLatched
 *   - SET:   runRequest=TRUE AND flameOK=FALSE  → same scan, no delay  [PUB001]
 *   - HOLD:  once set, retained across scans until valid reset edge     [PUB016]
 *   - RESET: rising(resetBtn) AND runRequest=FALSE AND flameOK=FALSE    [PUB016]
 *   - Edge-only reset; hold/rescan does NOT clear; press without edge does NOT clear
 * Output: fuelPermit
 *   - Activation:   runRequest AND flameOK AND NOT tripLatched          [PUB003]
 *   - Retention:    none — combinational, 0 when tripLatched           [PUB003]
 *   - Deactivation: tripLatched rising sets to FALSE; also 0 when any input low [PUB003]
 *   - Units: BOOLEAN
 * Output: trimEnable
 *   - Activation:   fuelPermit=TRUE AND o2Fault=FALSE                    [PUB008]
 *   - Retention:    none — combinational, 0 when o2Fault                [PUB008]
 *   - Deactivation: o2Fault rising (invalid/range)                      [PUB008]
 * Output: airTrim
 *   - Activation:   trimEnable with formula 2.0*(2.0-o2PV), clamp ±10   [PUB005]
 *   - Retention:    0.0 when trimEnable=FALSE (no residual)             [PUB010]
 *   - Units: % offset, clamped [-10,+10]
 * Output: airCommand
 *   - Activation:   baseAir+airTrim clamped [0,100] when fuelPermit=TRUE [PUB006]
 *   - Retention:    0.0 when fuelPermit=FALSE                           [PUB005]
 *   - Units: % absolute, clamped [0,100]; baseAir may be outside range [PUB006]
 * Output: o2Fault
 *   - Activation:   NOT o2Valid OR o2PV<0 OR o2PV>21                    [PUB009]
 *   - Retention:    combinational; does not inhibit fuelPermit          [PUB009]
 * Same-scan priority: trip set, fuelPermit, trimEnable/o2Fault, airTrim, airCommand
 * CONTRACT_RULES []
 *)
    // Detect rising edge of reset button (edge-only reset per PUB016)
    tmp_reset_rising := resetBtn AND NOT tmp_reset_rising;

    // Trip latch: set when running without flame, hold until valid reset edge
    tmp_trip_set := runRequest AND NOT flameOK;
    IF tmp_trip_set THEN
        tripLatched := TRUE;
    ELSIF tmp_reset_rising AND NOT runRequest AND NOT flameOK THEN
        tripLatched := FALSE;
    END_IF;

    // Fuel permit: requires run, flame, and no trip
    fuelPermit := runRequest AND flameOK AND NOT tripLatched;

    // O2 fault detection
    o2Fault := NOT o2Valid OR o2PV < 0.0 OR o2PV > 21.0;

    // Trim enable: fuel permit without O2 fault
    trimEnable := fuelPermit AND NOT o2Fault;

    // Air trim: 2.0*(2.0-o2PV), clamped to [-10, +10]; forced 0 when disabled
    IF trimEnable THEN
        airTrim := 2.0 * (2.0 - o2PV);
        IF airTrim > 10.0 THEN
            airTrim := 10.0;
        ELSIF airTrim < -10.0 THEN
            airTrim := -10.0;
        END_IF;
    ELSE
        airTrim := 0.0;
    END_IF;

    // Air command: base + trim, clamped [0,100]; forced 0 when no fuel permit
    IF fuelPermit THEN
        airCommand := baseAir + airTrim;
        IF airCommand > 100.0 THEN
            airCommand := 100.0;
        ELSIF airCommand < 0.0 THEN
            airCommand := 0.0;
        END_IF;
    ELSE
        airCommand := 0.0;
    END_IF;
END_FUNCTION_BLOCK

(* ---- self-hard-05.raw_candidate_01.st ---- *)
FUNCTION_BLOCK FB
VAR_INPUT
    runRequest  : BOOL;
    flameOK     : BOOL;
    o2Valid     : BOOL;
    o2PV        : REAL;
    baseAir     : REAL;
    resetBtn    : BOOL;
END_VAR
VAR_OUTPUT
    fuelPermit  : BOOL;
    trimEnable  : BOOL;
    airTrim     : REAL;
    airCommand  : REAL;
    tripLatched : BOOL;
    o2Fault     : BOOL;
END_VAR
VAR
    tmp_reset_rising : BOOL;
    tmp_trip_set     : BOOL;
END_VAR
(* ENGINEERING_CONTRACT
 * Output: tripLatched
 *   - SET:   runRequest=TRUE AND flameOK=FALSE  → same scan, no delay  [PUB001]
 *   - HOLD:  once set, retained across scans until valid reset edge     [PUB016]
 *   - RESET: rising(resetBtn) AND runRequest=FALSE AND flameOK=FALSE    [PUB016]
 *   - Edge-only reset; hold/rescan does NOT clear; press without edge does NOT clear
 * Output: fuelPermit
 *   - Activation:   runRequest AND flameOK AND NOT tripLatched          [PUB003]
 *   - Retention:    none — combinational, 0 when tripLatched           [PUB003]
 *   - Deactivation: tripLatched rising sets to FALSE; also 0 when any input low [PUB003]
 *   - Units: BOOLEAN
 * Output: trimEnable
 *   - Activation:   fuelPermit=TRUE AND o2Fault=FALSE                    [PUB008]
 *   - Retention:    none — combinational, 0 when o2Fault                [PUB008]
 *   - Deactivation: o2Fault rising (invalid/range)                      [PUB008]
 * Output: airTrim
 *   - Activation:   trimEnable with formula 2.0*(2.0-o2PV), clamp ±10   [PUB005]
 *   - Retention:    0.0 when trimEnable=FALSE (no residual)             [PUB010]
 *   - Units: % offset, clamped [-10,+10]
 * Output: airCommand
 *   - Activation:   baseAir+airTrim clamped [0,100] when fuelPermit=TRUE [PUB006]
 *   - Retention:    0.0 when fuelPermit=FALSE                           [PUB005]
 *   - Units: % absolute, clamped [0,100]; baseAir may be outside range [PUB006]
 * Output: o2Fault
 *   - Activation:   NOT o2Valid OR o2PV<0 OR o2PV>21                    [PUB009]
 *   - Retention:    combinational; does not inhibit fuelPermit          [PUB009]
 * Same-scan priority: trip set, fuelPermit, trimEnable/o2Fault, airTrim, airCommand
 * CONTRACT_RULES []
 *)
    // Detect rising edge of reset button (edge-only reset per PUB016)
    tmp_reset_rising := resetBtn AND NOT tmp_reset_rising;

    // Trip latch: set when running without flame, hold until valid reset edge
    tmp_trip_set := runRequest AND NOT flameOK;
    IF tmp_trip_set THEN
        tripLatched := TRUE;
    ELSIF tmp_reset_rising AND NOT runRequest AND NOT flameOK THEN
        tripLatched := FALSE;
    END_IF;

    // Fuel permit: requires run, flame, and no trip
    fuelPermit := runRequest AND flameOK AND NOT tripLatched;

    // O2 fault detection
    o2Fault := NOT o2Valid OR o2PV < 0.0 OR o2PV > 21.0;

    // Trim enable: fuel permit without O2 fault
    trimEnable := fuelPermit AND NOT o2Fault;

    // Air trim: 2.0*(2.0-o2PV), clamped to [-10, +10]; forced 0 when disabled
    IF trimEnable THEN
        airTrim := 2.0 * (2.0 - o2PV);
        IF airTrim > 10.0 THEN
            airTrim := 10.0;
        ELSIF airTrim < -10.0 THEN
            airTrim := -10.0;
        END_IF;
    ELSE
        airTrim := 0.0;
    END_IF;

    // Air command: base + trim, clamped [0,100]; forced 0 when no fuel permit
    IF fuelPermit THEN
        airCommand := baseAir + airTrim;
        IF airCommand > 100.0 THEN
            airCommand := 100.0;
        ELSIF airCommand < 0.0 THEN
            airCommand := 0.0;
        END_IF;
    ELSE
        airCommand := 0.0;
    END_IF;
END_FUNCTION_BLOCK

(* ---- self-hard-06.candidate_01.st ---- *)
(* ENGINEERING_CONTRACT: Steam Header Overpressure Interlock + Fault Diagnosis
 * ================================================================================
 * [PUB001] Function: FB - steam header overpressure interlock with fault footprint
 * [PUB002] Trip activation: runRequest AND (NOT pressureValid OR pressure >= 4500.0) same-scan
 * [PUB003] Reset permission: resetBtn rising-edge AND NOT runRequest AND pressureValid AND pressure <= 4200.0
 * [PUB004] Hysteresis: 300 kPa (4500 trip / 4200 reset gap per PUB003/PUB010)
 * [PUB005] Fault bit0=1: runRequest AND NOT pressureValid (transmitter failure)
 * [PUB006] Fault bit1=2: outletCmd>=50 AND outletFeedback<=10 for 3 consecutive valid overpressure scans
 *            Counter reset on: NOT runRequest, NOT pressureValid, pressure<4500, or condition unsatisfied
 * [PUB007] Fault bit2=4: fuelFlow >= 4.0 AND steamFlow <= 10.0 (valid overpressure工况 only)
 * [PUB008] Fault bit3=8: overpressure but no specific cause identified (valid overpressure工况 only)
 * [PUB009] currentCauseMask reset to 0 when NOT runRequest; low 4 bits only; allowed: 0,1,2,4,6,8
 * [PUB010] latchedCauseMask: bitwise OR accumulation while tripLatched=TRUE; cleared on valid reset only
 * [PUB011] fuelPermit = runRequest AND NOT tripLatched; diagnosticActive = currentCauseMask <> 0
 * [PUB012] Output retention: tripLatched holds until valid reset; fuelPermit combinational per PUB011
 * [PUB013] Units: kPa (pressure), t/h (flow), % (valve), dimensionless (bit masks)
 * [PUB014] No hidden timers; all state in VAR; same-scan evaluation per PUB002
 *
 * CONTRACT_RULES [{"kind":"hold_until_reset","output":"tripLatched","set_input":"runRequest","reset_input":"resetBtn"}]
 *)
FUNCTION_BLOCK FB
VAR_INPUT
    runRequest      : BOOL;
    pressure        : REAL;
    pressureValid   : BOOL;
    fuelFlow        : REAL;
    steamFlow       : REAL;
    outletCmd       : INT;
    outletFeedback  : INT;
    resetBtn        : BOOL;
END_VAR
VAR_OUTPUT
    tripLatched     : BOOL;
    fuelPermit      : BOOL;
    currentCauseMask: WORD;
    latchedCauseMask: WORD;
    diagnosticActive: BOOL;
END_VAR
VAR
    prevResetBtn    : BOOL := FALSE;
    prevRunRequest  : BOOL := FALSE;
    stuckCnt        : INT  := 0;
END_VAR

// ---- Rising-edge detection for reset button ----
IF resetBtn AND NOT prevResetBtn THEN
    // Rising edge of resetBtn
    IF NOT runRequest AND pressureValid AND pressure <= 4200.0 THEN
        tripLatched     := FALSE;
        latchedCauseMask := 0;
    END_IF;
END_IF;
prevResetBtn := resetBtn;

// ---- Trip latch activation (PUB002) ----
IF runRequest AND (NOT pressureValid OR pressure >= 4500.0) THEN
    tripLatched := TRUE;
END_IF;

// ---- Fault diagnosis: currentCauseMask (PUB005-PUB009) ----
VAR tempMask : WORD := 0; END_VAR
// bit0: transmitter failure (overrides all other conditions per PUB012)
IF runRequest AND NOT pressureValid THEN
    tempMask := 1; // bit0=1
ELSE
    // bit1 and bit2 only evaluated in valid overpressure工况 (PUB008/PUB009)
    IF runRequest AND pressureValid AND pressure >= 4500.0 THEN
        // Stuck valve counter: 3 consecutive valid scans (PUB006)
        IF outletCmd >= 50 AND outletFeedback <= 10 THEN
            stuckCnt := stuckCnt + 1;
        ELSE
            stuckCnt := 0;
        END_IF;
        IF stuckCnt >= 3 THEN
            tempMask := tempMask OR 2; // bit1=2
        END_IF;
        // Excess combustion: fuelFlow>=4.0 AND steamFlow<=10.0 (PUB007)
        IF fuelFlow >= 4.0 AND steamFlow <= 10.0 THEN
            tempMask := tempMask OR 4; // bit2=4
        END_IF;
        // Unlocated: overpressure but no specific cause (PUB008)
        IF tempMask = 0 THEN
            tempMask := 8; // bit3=8
        END_IF;
    ELSE
        stuckCnt := 0;
    END_IF;
ELSE
    stuckCnt := 0;
END_IF;
currentCauseMask := tempMask;

// ---- Latched cause accumulation (PUB010) ----
IF tripLatched THEN
    latchedCauseMask := latchedCauseMask OR currentCauseMask;
END_IF;

// ---- Fuel permit and diagnostic (PUB011) ----
fuelPermit      := runRequest AND NOT tripLatched;
diagnosticActive := currentCauseMask <> 0;

// ---- Update previous run state for rising-edge tracking ----
prevRunRequest := runRequest;
END_FUNCTION_BLOCK

(* ---- self-hard-06.candidate_02.st ---- *)
(* ENGINEERING_CONTRACT: Steam Header Overpressure Interlock + Fault Diagnosis
 * ================================================================================
 * [PUB001] Function: FB - steam header overpressure interlock with fault footprint
 * [PUB002] Trip activation: runRequest AND (NOT pressureValid OR pressure >= 4500.0) same-scan
 * [PUB003] Reset permission: resetBtn rising-edge AND NOT runRequest AND pressureValid AND pressure <= 4200.0
 * [PUB004] Hysteresis: 300 kPa (4500 trip / 4200 reset gap per PUB003/PUB010)
 * [PUB005] Fault bit0=1: runRequest AND NOT pressureValid (transmitter failure)
 * [PUB006] Fault bit1=2: outletCmd>=50 AND outletFeedback<=10 for 3 consecutive valid overpressure scans
 *            Counter reset on: NOT runRequest, NOT pressureValid, pressure<4500, or condition unsatisfied
 * [PUB007] Fault bit2=4: fuelFlow >= 4.0 AND steamFlow <= 10.0 (valid overpressure工况 only)
 * [PUB008] Fault bit3=8: overpressure but no specific cause identified (valid overpressure工况 only)
 * [PUB009] currentCauseMask reset to 0 when NOT runRequest; low 4 bits only; allowed: 0,1,2,4,6,8
 * [PUB010] latchedCauseMask: bitwise OR accumulation while tripLatched=TRUE; cleared on valid reset only
 * [PUB011] fuelPermit = runRequest AND NOT tripLatched; diagnosticActive = currentCauseMask <> 0
 * [PUB012] Output retention: tripLatched holds until valid reset; fuelPermit combinational per PUB011
 * [PUB013] Units: kPa (pressure), t/h (flow), % (valve), dimensionless (bit masks)
 * [PUB014] No hidden timers; all state in VAR; same-scan evaluation per PUB002
 *
 * CONTRACT_RULES [{"kind":"hold_until_reset","output":"tripLatched","set_input":"runRequest","reset_input":"resetBtn"}]
 *)
FUNCTION_BLOCK FB
VAR_INPUT
    runRequest      : BOOL;
    pressure        : REAL;
    pressureValid   : BOOL;
    fuelFlow        : REAL;
    steamFlow       : REAL;
    outletCmd       : INT;
    outletFeedback  : INT;
    resetBtn        : BOOL;
END_VAR
VAR_OUTPUT
    tripLatched     : BOOL;
    fuelPermit      : BOOL;
    currentCauseMask: WORD;
    latchedCauseMask: WORD;
    diagnosticActive: BOOL;
END_VAR
VAR
    prevResetBtn    : BOOL := FALSE;
    prevRunRequest  : BOOL := FALSE;
    stuckCnt        : INT  := 0;
    tempMask        : WORD := 0;
END_VAR

// ---- Rising-edge detection for reset button ----
IF resetBtn AND NOT prevResetBtn THEN
    // Rising edge of resetBtn
    IF NOT runRequest AND pressureValid AND pressure <= 4200.0 THEN
        tripLatched     := FALSE;
        latchedCauseMask := 0;
    END_IF;
END_IF;
prevResetBtn := resetBtn;

// ---- Trip latch activation (PUB002) ----
IF runRequest AND (NOT pressureValid OR pressure >= 4500.0) THEN
    tripLatched := TRUE;
END_IF;

// ---- Fault diagnosis: currentCauseMask (PUB005-PUB009) ----
VAR tempMask : WORD := 0; END_VAR
// bit0: transmitter failure (overrides all other conditions per PUB012)
IF runRequest AND NOT pressureValid THEN
    tempMask := 1; // bit0=1
ELSE
    // bit1 and bit2 only evaluated in valid overpressure工况 (PUB008/PUB009)
    IF runRequest AND pressureValid AND pressure >= 4500.0 THEN
        // Stuck valve counter: 3 consecutive valid scans (PUB006)
        IF outletCmd >= 50 AND outletFeedback <= 10 THEN
            stuckCnt := stuckCnt + 1;
        ELSE
            stuckCnt := 0;
        END_IF;
        IF stuckCnt >= 3 THEN
            tempMask := tempMask OR 2; // bit1=2
        END_IF;
        // Excess combustion: fuelFlow>=4.0 AND steamFlow<=10.0 (PUB007)
        IF fuelFlow >= 4.0 AND steamFlow <= 10.0 THEN
            tempMask := tempMask OR 4; // bit2=4
        END_IF;
        // Unlocated: overpressure but no specific cause (PUB008)
        IF tempMask = 0 THEN
            tempMask := 8; // bit3=8
        END_IF;
    ELSE
        stuckCnt := 0;
    END_IF;
ELSE
    stuckCnt := 0;
END_IF;
currentCauseMask := tempMask;

// ---- Latched cause accumulation (PUB010) ----
IF tripLatched THEN
    latchedCauseMask := latchedCauseMask OR currentCauseMask;
END_IF;

// ---- Fuel permit and diagnostic (PUB011) ----
fuelPermit      := runRequest AND NOT tripLatched;
diagnosticActive := currentCauseMask <> 0;

// ---- Update previous run state for rising-edge tracking ----
prevRunRequest := runRequest;
END_FUNCTION_BLOCK

(* ---- self-hard-06.candidate_03.st ---- *)
(* ENGINEERING_CONTRACT: Steam Header Overpressure Interlock + Fault Diagnosis
 * ================================================================================
 * [PUB001] Function: FB - steam header overpressure interlock with fault footprint
 * [PUB002] Trip activation: runRequest AND (NOT pressureValid OR pressure >= 4500.0) same-scan
 * [PUB003] Reset permission: resetBtn rising-edge AND NOT runRequest AND pressureValid AND pressure <= 4200.0
 * [PUB004] Hysteresis: 300 kPa (4500 trip / 4200 reset gap per PUB003/PUB010)
 * [PUB005] Fault bit0=1: runRequest AND NOT pressureValid (transmitter failure)
 * [PUB006] Fault bit1=2: outletCmd>=50 AND outletFeedback<=10 for 3 consecutive valid overpressure scans
 *            Counter reset on: NOT runRequest, NOT pressureValid, pressure<4500, or condition unsatisfied
 * [PUB007] Fault bit2=4: fuelFlow >= 4.0 AND steamFlow <= 10.0 (valid overpressure工况 only)
 * [PUB008] Fault bit3=8: overpressure but no specific cause identified (valid overpressure工况 only)
 * [PUB009] currentCauseMask reset to 0 when NOT runRequest; low 4 bits only; allowed: 0,1,2,4,6,8
 * [PUB010] latchedCauseMask: bitwise OR accumulation while tripLatched=TRUE; cleared on valid reset only
 * [PUB011] fuelPermit = runRequest AND NOT tripLatched; diagnosticActive = currentCauseMask <> 0
 * [PUB012] Output retention: tripLatched holds until valid reset; fuelPermit combinational per PUB011
 * [PUB013] Units: kPa (pressure), t/h (flow), % (valve), dimensionless (bit masks)
 * [PUB014] No hidden timers; all state in VAR; same-scan evaluation per PUB002
 *
 * CONTRACT_RULES [{"kind":"hold_until_reset","output":"tripLatched","set_input":"runRequest","reset_input":"resetBtn"}]
 *)
FUNCTION_BLOCK FB
VAR_INPUT
    runRequest      : BOOL;
    pressure        : REAL;
    pressureValid   : BOOL;
    fuelFlow        : REAL;
    steamFlow       : REAL;
    outletCmd       : INT;
    outletFeedback  : INT;
    resetBtn        : BOOL;
END_VAR
VAR_OUTPUT
    tripLatched     : BOOL;
    fuelPermit      : BOOL;
    currentCauseMask: WORD;
    latchedCauseMask: WORD;
    diagnosticActive: BOOL;
END_VAR
VAR
    prevResetBtn    : BOOL := FALSE;
    prevRunRequest  : BOOL := FALSE;
    stuckCnt        : INT  := 0;
    tempMask        : WORD := 0;
END_VAR

// ---- Rising-edge detection for reset button ----
IF resetBtn AND NOT prevResetBtn THEN
    IF NOT runRequest AND pressureValid AND pressure <= 4200.0 THEN
        tripLatched      := FALSE;
        latchedCauseMask := 0;
    END_IF;
END_IF;
prevResetBtn := resetBtn;

// ---- Trip latch activation (PUB002) ----
IF runRequest AND (NOT pressureValid OR pressure >= 4500.0) THEN
    tripLatched := TRUE;
END_IF;

// ---- Fault diagnosis: currentCauseMask (PUB005-PUB009) ----
tempMask := 0;
IF runRequest AND NOT pressureValid THEN
    tempMask := 1;
ELSIF runRequest AND pressureValid AND pressure >= 4500.0 THEN
    IF outletCmd >= 50 AND outletFeedback <= 10 THEN
        stuckCnt := stuckCnt + 1;
    ELSE
        stuckCnt := 0;
    END_IF;
    IF stuckCnt >= 3 THEN
        tempMask := tempMask OR 2;
    END_IF;
    IF fuelFlow >= 4.0 AND steamFlow <= 10.0 THEN
        tempMask := tempMask OR 4;
    END_IF;
    IF tempMask = 0 THEN
        tempMask := 8;
    END_IF;
ELSE
    stuckCnt := 0;
END_IF;
currentCauseMask := tempMask;

// ---- Latched cause accumulation (PUB010) ----
IF tripLatched THEN
    latchedCauseMask := latchedCauseMask OR currentCauseMask;
END_IF;

// ---- Fuel permit and diagnostic (PUB011) ----
fuelPermit      := runRequest AND NOT tripLatched;
diagnosticActive := currentCauseMask <> 0;

// ---- Update previous run state for rising-edge tracking ----
prevRunRequest := runRequest;
END_FUNCTION_BLOCK

(* ---- self-hard-06.patch_base_02.st ---- *)
(* ENGINEERING_CONTRACT: Steam Header Overpressure Interlock + Fault Diagnosis
 * ================================================================================
 * [PUB001] Function: FB - steam header overpressure interlock with fault footprint
 * [PUB002] Trip activation: runRequest AND (NOT pressureValid OR pressure >= 4500.0) same-scan
 * [PUB003] Reset permission: resetBtn rising-edge AND NOT runRequest AND pressureValid AND pressure <= 4200.0
 * [PUB004] Hysteresis: 300 kPa (4500 trip / 4200 reset gap per PUB003/PUB010)
 * [PUB005] Fault bit0=1: runRequest AND NOT pressureValid (transmitter failure)
 * [PUB006] Fault bit1=2: outletCmd>=50 AND outletFeedback<=10 for 3 consecutive valid overpressure scans
 *            Counter reset on: NOT runRequest, NOT pressureValid, pressure<4500, or condition unsatisfied
 * [PUB007] Fault bit2=4: fuelFlow >= 4.0 AND steamFlow <= 10.0 (valid overpressure工况 only)
 * [PUB008] Fault bit3=8: overpressure but no specific cause identified (valid overpressure工况 only)
 * [PUB009] currentCauseMask reset to 0 when NOT runRequest; low 4 bits only; allowed: 0,1,2,4,6,8
 * [PUB010] latchedCauseMask: bitwise OR accumulation while tripLatched=TRUE; cleared on valid reset only
 * [PUB011] fuelPermit = runRequest AND NOT tripLatched; diagnosticActive = currentCauseMask <> 0
 * [PUB012] Output retention: tripLatched holds until valid reset; fuelPermit combinational per PUB011
 * [PUB013] Units: kPa (pressure), t/h (flow), % (valve), dimensionless (bit masks)
 * [PUB014] No hidden timers; all state in VAR; same-scan evaluation per PUB002
 *
 * CONTRACT_RULES [{"kind":"hold_until_reset","output":"tripLatched","set_input":"runRequest","reset_input":"resetBtn"}]
 *)
FUNCTION_BLOCK FB
VAR_INPUT
    runRequest      : BOOL;
    pressure        : REAL;
    pressureValid   : BOOL;
    fuelFlow        : REAL;
    steamFlow       : REAL;
    outletCmd       : INT;
    outletFeedback  : INT;
    resetBtn        : BOOL;
END_VAR
VAR_OUTPUT
    tripLatched     : BOOL;
    fuelPermit      : BOOL;
    currentCauseMask: WORD;
    latchedCauseMask: WORD;
    diagnosticActive: BOOL;
END_VAR
VAR
    prevResetBtn    : BOOL := FALSE;
    prevRunRequest  : BOOL := FALSE;
    stuckCnt        : INT  := 0;
END_VAR

// ---- Rising-edge detection for reset button ----
IF resetBtn AND NOT prevResetBtn THEN
    // Rising edge of resetBtn
    IF NOT runRequest AND pressureValid AND pressure <= 4200.0 THEN
        tripLatched     := FALSE;
        latchedCauseMask := 0;
    END_IF;
END_IF;
prevResetBtn := resetBtn;

// ---- Trip latch activation (PUB002) ----
IF runRequest AND (NOT pressureValid OR pressure >= 4500.0) THEN
    tripLatched := TRUE;
END_IF;

// ---- Fault diagnosis: currentCauseMask (PUB005-PUB009) ----
VAR tempMask : WORD := 0; END_VAR
// bit0: transmitter failure (overrides all other conditions per PUB012)
IF runRequest AND NOT pressureValid THEN
    tempMask := 1; // bit0=1
ELSE
    // bit1 and bit2 only evaluated in valid overpressure工况 (PUB008/PUB009)
    IF runRequest AND pressureValid AND pressure >= 4500.0 THEN
        // Stuck valve counter: 3 consecutive valid scans (PUB006)
        IF outletCmd >= 50 AND outletFeedback <= 10 THEN
            stuckCnt := stuckCnt + 1;
        ELSE
            stuckCnt := 0;
        END_IF;
        IF stuckCnt >= 3 THEN
            tempMask := tempMask OR 2; // bit1=2
        END_IF;
        // Excess combustion: fuelFlow>=4.0 AND steamFlow<=10.0 (PUB007)
        IF fuelFlow >= 4.0 AND steamFlow <= 10.0 THEN
            tempMask := tempMask OR 4; // bit2=4
        END_IF;
        // Unlocated: overpressure but no specific cause (PUB008)
        IF tempMask = 0 THEN
            tempMask := 8; // bit3=8
        END_IF;
    ELSE
        stuckCnt := 0;
    END_IF;
ELSE
    stuckCnt := 0;
END_IF;
currentCauseMask := tempMask;

// ---- Latched cause accumulation (PUB010) ----
IF tripLatched THEN
    latchedCauseMask := latchedCauseMask OR currentCauseMask;
END_IF;

// ---- Fuel permit and diagnostic (PUB011) ----
fuelPermit      := runRequest AND NOT tripLatched;
diagnosticActive := currentCauseMask <> 0;

// ---- Update previous run state for rising-edge tracking ----
prevRunRequest := runRequest;
END_FUNCTION_BLOCK

(* ---- self-hard-06.patch_base_03.st ---- *)
(* ENGINEERING_CONTRACT: Steam Header Overpressure Interlock + Fault Diagnosis
 * ================================================================================
 * [PUB001] Function: FB - steam header overpressure interlock with fault footprint
 * [PUB002] Trip activation: runRequest AND (NOT pressureValid OR pressure >= 4500.0) same-scan
 * [PUB003] Reset permission: resetBtn rising-edge AND NOT runRequest AND pressureValid AND pressure <= 4200.0
 * [PUB004] Hysteresis: 300 kPa (4500 trip / 4200 reset gap per PUB003/PUB010)
 * [PUB005] Fault bit0=1: runRequest AND NOT pressureValid (transmitter failure)
 * [PUB006] Fault bit1=2: outletCmd>=50 AND outletFeedback<=10 for 3 consecutive valid overpressure scans
 *            Counter reset on: NOT runRequest, NOT pressureValid, pressure<4500, or condition unsatisfied
 * [PUB007] Fault bit2=4: fuelFlow >= 4.0 AND steamFlow <= 10.0 (valid overpressure工况 only)
 * [PUB008] Fault bit3=8: overpressure but no specific cause identified (valid overpressure工况 only)
 * [PUB009] currentCauseMask reset to 0 when NOT runRequest; low 4 bits only; allowed: 0,1,2,4,6,8
 * [PUB010] latchedCauseMask: bitwise OR accumulation while tripLatched=TRUE; cleared on valid reset only
 * [PUB011] fuelPermit = runRequest AND NOT tripLatched; diagnosticActive = currentCauseMask <> 0
 * [PUB012] Output retention: tripLatched holds until valid reset; fuelPermit combinational per PUB011
 * [PUB013] Units: kPa (pressure), t/h (flow), % (valve), dimensionless (bit masks)
 * [PUB014] No hidden timers; all state in VAR; same-scan evaluation per PUB002
 *
 * CONTRACT_RULES [{"kind":"hold_until_reset","output":"tripLatched","set_input":"runRequest","reset_input":"resetBtn"}]
 *)
FUNCTION_BLOCK FB
VAR_INPUT
    runRequest      : BOOL;
    pressure        : REAL;
    pressureValid   : BOOL;
    fuelFlow        : REAL;
    steamFlow       : REAL;
    outletCmd       : INT;
    outletFeedback  : INT;
    resetBtn        : BOOL;
END_VAR
VAR_OUTPUT
    tripLatched     : BOOL;
    fuelPermit      : BOOL;
    currentCauseMask: WORD;
    latchedCauseMask: WORD;
    diagnosticActive: BOOL;
END_VAR
VAR
    prevResetBtn    : BOOL := FALSE;
    prevRunRequest  : BOOL := FALSE;
    stuckCnt        : INT  := 0;
END_VAR

// ---- Rising-edge detection for reset button ----
IF resetBtn AND NOT prevResetBtn THEN
    // Rising edge of resetBtn
    IF NOT runRequest AND pressureValid AND pressure <= 4200.0 THEN
        tripLatched     := FALSE;
        latchedCauseMask := 0;
    END_IF;
END_IF;
prevResetBtn := resetBtn;

// ---- Trip latch activation (PUB002) ----
IF runRequest AND (NOT pressureValid OR pressure >= 4500.0) THEN
    tripLatched := TRUE;
END_IF;

// ---- Fault diagnosis: currentCauseMask (PUB005-PUB009) ----
VAR tempMask : WORD := 0; END_VAR
// bit0: transmitter failure (overrides all other conditions per PUB012)
IF runRequest AND NOT pressureValid THEN
    tempMask := 1; // bit0=1
ELSE
    // bit1 and bit2 only evaluated in valid overpressure工况 (PUB008/PUB009)
    IF runRequest AND pressureValid AND pressure >= 4500.0 THEN
        // Stuck valve counter: 3 consecutive valid scans (PUB006)
        IF outletCmd >= 50 AND outletFeedback <= 10 THEN
            stuckCnt := stuckCnt + 1;
        ELSE
            stuckCnt := 0;
        END_IF;
        IF stuckCnt >= 3 THEN
            tempMask := tempMask OR 2; // bit1=2
        END_IF;
        // Excess combustion: fuelFlow>=4.0 AND steamFlow<=10.0 (PUB007)
        IF fuelFlow >= 4.0 AND steamFlow <= 10.0 THEN
            tempMask := tempMask OR 4; // bit2=4
        END_IF;
        // Unlocated: overpressure but no specific cause (PUB008)
        IF tempMask = 0 THEN
            tempMask := 8; // bit3=8
        END_IF;
    ELSE
        stuckCnt := 0;
    END_IF;
ELSE
    stuckCnt := 0;
END_IF;
currentCauseMask := tempMask;

// ---- Latched cause accumulation (PUB010) ----
IF tripLatched THEN
    latchedCauseMask := latchedCauseMask OR currentCauseMask;
END_IF;

// ---- Fuel permit and diagnostic (PUB011) ----
fuelPermit      := runRequest AND NOT tripLatched;
diagnosticActive := currentCauseMask <> 0;

// ---- Update previous run state for rising-edge tracking ----
prevRunRequest := runRequest;
END_FUNCTION_BLOCK

(* ---- self-hard-06.patch_base_04.st ---- *)
(* ENGINEERING_CONTRACT: Steam Header Overpressure Interlock + Fault Diagnosis
 * ================================================================================
 * [PUB001] Function: FB - steam header overpressure interlock with fault footprint
 * [PUB002] Trip activation: runRequest AND (NOT pressureValid OR pressure >= 4500.0) same-scan
 * [PUB003] Reset permission: resetBtn rising-edge AND NOT runRequest AND pressureValid AND pressure <= 4200.0
 * [PUB004] Hysteresis: 300 kPa (4500 trip / 4200 reset gap per PUB003/PUB010)
 * [PUB005] Fault bit0=1: runRequest AND NOT pressureValid (transmitter failure)
 * [PUB006] Fault bit1=2: outletCmd>=50 AND outletFeedback<=10 for 3 consecutive valid overpressure scans
 *            Counter reset on: NOT runRequest, NOT pressureValid, pressure<4500, or condition unsatisfied
 * [PUB007] Fault bit2=4: fuelFlow >= 4.0 AND steamFlow <= 10.0 (valid overpressure工况 only)
 * [PUB008] Fault bit3=8: overpressure but no specific cause identified (valid overpressure工况 only)
 * [PUB009] currentCauseMask reset to 0 when NOT runRequest; low 4 bits only; allowed: 0,1,2,4,6,8
 * [PUB010] latchedCauseMask: bitwise OR accumulation while tripLatched=TRUE; cleared on valid reset only
 * [PUB011] fuelPermit = runRequest AND NOT tripLatched; diagnosticActive = currentCauseMask <> 0
 * [PUB012] Output retention: tripLatched holds until valid reset; fuelPermit combinational per PUB011
 * [PUB013] Units: kPa (pressure), t/h (flow), % (valve), dimensionless (bit masks)
 * [PUB014] No hidden timers; all state in VAR; same-scan evaluation per PUB002
 *
 * CONTRACT_RULES [{"kind":"hold_until_reset","output":"tripLatched","set_input":"runRequest","reset_input":"resetBtn"}]
 *)
FUNCTION_BLOCK FB
VAR_INPUT
    runRequest      : BOOL;
    pressure        : REAL;
    pressureValid   : BOOL;
    fuelFlow        : REAL;
    steamFlow       : REAL;
    outletCmd       : INT;
    outletFeedback  : INT;
    resetBtn        : BOOL;
END_VAR
VAR_OUTPUT
    tripLatched     : BOOL;
    fuelPermit      : BOOL;
    currentCauseMask: WORD;
    latchedCauseMask: WORD;
    diagnosticActive: BOOL;
END_VAR
VAR
    prevResetBtn    : BOOL := FALSE;
    prevRunRequest  : BOOL := FALSE;
    stuckCnt        : INT  := 0;
    tempMask        : WORD := 0;
END_VAR

// ---- Rising-edge detection for reset button ----
IF resetBtn AND NOT prevResetBtn THEN
    IF NOT runRequest AND pressureValid AND pressure <= 4200.0 THEN
        tripLatched      := FALSE;
        latchedCauseMask := 0;
    END_IF;
END_IF;
prevResetBtn := resetBtn;

// ---- Trip latch activation (PUB002) ----
IF runRequest AND (NOT pressureValid OR pressure >= 4500.0) THEN
    tripLatched := TRUE;
END_IF;

// ---- Fault diagnosis: currentCauseMask (PUB005-PUB009) ----
tempMask := 0;
IF runRequest AND NOT pressureValid THEN
    tempMask := 1;
ELSIF runRequest AND pressureValid AND pressure >= 4500.0 THEN
    IF outletCmd >= 50 AND outletFeedback <= 10 THEN
        stuckCnt := stuckCnt + 1;
    ELSE
        stuckCnt := 0;
    END_IF;
    IF stuckCnt >= 3 THEN
        tempMask := tempMask OR 2;
    END_IF;
    IF fuelFlow >= 4.0 AND steamFlow <= 10.0 THEN
        tempMask := tempMask OR 4;
    END_IF;
    IF tempMask = 0 THEN
        tempMask := 8;
    END_IF;
ELSE
    stuckCnt := 0;
END_IF;
currentCauseMask := tempMask;

// ---- Latched cause accumulation (PUB010) ----
IF tripLatched THEN
    latchedCauseMask := latchedCauseMask OR currentCauseMask;
END_IF;

// ---- Fuel permit and diagnostic (PUB011) ----
fuelPermit      := runRequest AND NOT tripLatched;
diagnosticActive := currentCauseMask <> 0;

// ---- Update previous run state for rising-edge tracking ----
prevRunRequest := runRequest;
END_FUNCTION_BLOCK

(* ---- self-hard-06.raw_candidate_01.st ---- *)
(* ENGINEERING_CONTRACT: Steam Header Overpressure Interlock + Fault Diagnosis
 * ================================================================================
 * [PUB001] Function: FB - steam header overpressure interlock with fault footprint
 * [PUB002] Trip activation: runRequest AND (NOT pressureValid OR pressure >= 4500.0) same-scan
 * [PUB003] Reset permission: resetBtn rising-edge AND NOT runRequest AND pressureValid AND pressure <= 4200.0
 * [PUB004] Hysteresis: 300 kPa (4500 trip / 4200 reset gap per PUB003/PUB010)
 * [PUB005] Fault bit0=1: runRequest AND NOT pressureValid (transmitter failure)
 * [PUB006] Fault bit1=2: outletCmd>=50 AND outletFeedback<=10 for 3 consecutive valid overpressure scans
 *            Counter reset on: NOT runRequest, NOT pressureValid, pressure<4500, or condition unsatisfied
 * [PUB007] Fault bit2=4: fuelFlow >= 4.0 AND steamFlow <= 10.0 (valid overpressure工况 only)
 * [PUB008] Fault bit3=8: overpressure but no specific cause identified (valid overpressure工况 only)
 * [PUB009] currentCauseMask reset to 0 when NOT runRequest; low 4 bits only; allowed: 0,1,2,4,6,8
 * [PUB010] latchedCauseMask: bitwise OR accumulation while tripLatched=TRUE; cleared on valid reset only
 * [PUB011] fuelPermit = runRequest AND NOT tripLatched; diagnosticActive = currentCauseMask <> 0
 * [PUB012] Output retention: tripLatched holds until valid reset; fuelPermit combinational per PUB011
 * [PUB013] Units: kPa (pressure), t/h (flow), % (valve), dimensionless (bit masks)
 * [PUB014] No hidden timers; all state in VAR; same-scan evaluation per PUB002
 *
 * CONTRACT_RULES [{"kind":"hold_until_reset","output":"tripLatched","set_input":"runRequest","reset_input":"resetBtn"}]
 *)
FUNCTION_BLOCK FB
VAR_INPUT
    runRequest      : BOOL;
    pressure        : REAL;
    pressureValid   : BOOL;
    fuelFlow        : REAL;
    steamFlow       : REAL;
    outletCmd       : INT;
    outletFeedback  : INT;
    resetBtn        : BOOL;
END_VAR
VAR_OUTPUT
    tripLatched     : BOOL;
    fuelPermit      : BOOL;
    currentCauseMask: WORD;
    latchedCauseMask: WORD;
    diagnosticActive: BOOL;
END_VAR
VAR
    prevResetBtn    : BOOL := FALSE;
    prevRunRequest  : BOOL := FALSE;
    stuckCnt        : INT  := 0;
END_VAR

// ---- Rising-edge detection for reset button ----
IF resetBtn AND NOT prevResetBtn THEN
    // Rising edge of resetBtn
    IF NOT runRequest AND pressureValid AND pressure <= 4200.0 THEN
        tripLatched     := FALSE;
        latchedCauseMask := 0;
    END_IF;
END_IF;
prevResetBtn := resetBtn;

// ---- Trip latch activation (PUB002) ----
IF runRequest AND (NOT pressureValid OR pressure >= 4500.0) THEN
    tripLatched := TRUE;
END_IF;

// ---- Fault diagnosis: currentCauseMask (PUB005-PUB009) ----
VAR tempMask : WORD := 0; END_VAR
// bit0: transmitter failure (overrides all other conditions per PUB012)
IF runRequest AND NOT pressureValid THEN
    tempMask := 1; // bit0=1
ELSE
    // bit1 and bit2 only evaluated in valid overpressure工况 (PUB008/PUB009)
    IF runRequest AND pressureValid AND pressure >= 4500.0 THEN
        // Stuck valve counter: 3 consecutive valid scans (PUB006)
        IF outletCmd >= 50 AND outletFeedback <= 10 THEN
            stuckCnt := stuckCnt + 1;
        ELSE
            stuckCnt := 0;
        END_IF;
        IF stuckCnt >= 3 THEN
            tempMask := tempMask OR 2; // bit1=2
        END_IF;
        // Excess combustion: fuelFlow>=4.0 AND steamFlow<=10.0 (PUB007)
        IF fuelFlow >= 4.0 AND steamFlow <= 10.0 THEN
            tempMask := tempMask OR 4; // bit2=4
        END_IF;
        // Unlocated: overpressure but no specific cause (PUB008)
        IF tempMask = 0 THEN
            tempMask := 8; // bit3=8
        END_IF;
    ELSE
        stuckCnt := 0;
    END_IF;
ELSE
    stuckCnt := 0;
END_IF;
currentCauseMask := tempMask;

// ---- Latched cause accumulation (PUB010) ----
IF tripLatched THEN
    latchedCauseMask := latchedCauseMask OR currentCauseMask;
END_IF;

// ---- Fuel permit and diagnostic (PUB011) ----
fuelPermit      := runRequest AND NOT tripLatched;
diagnosticActive := currentCauseMask <> 0;

// ---- Update previous run state for rising-edge tracking ----
prevRunRequest := runRequest;
END_FUNCTION_BLOCK

(* ---- self-hard-06.raw_candidate_02.st ---- *)
(* ENGINEERING_CONTRACT: Steam Header Overpressure Interlock + Fault Diagnosis
 * ================================================================================
 * [PUB001] Function: FB - steam header overpressure interlock with fault footprint
 * [PUB002] Trip activation: runRequest AND (NOT pressureValid OR pressure >= 4500.0) same-scan
 * [PUB003] Reset permission: resetBtn rising-edge AND NOT runRequest AND pressureValid AND pressure <= 4200.0
 * [PUB004] Hysteresis: 300 kPa (4500 trip / 4200 reset gap per PUB003/PUB010)
 * [PUB005] Fault bit0=1: runRequest AND NOT pressureValid (transmitter failure)
 * [PUB006] Fault bit1=2: outletCmd>=50 AND outletFeedback<=10 for 3 consecutive valid overpressure scans
 *            Counter reset on: NOT runRequest, NOT pressureValid, pressure<4500, or condition unsatisfied
 * [PUB007] Fault bit2=4: fuelFlow >= 4.0 AND steamFlow <= 10.0 (valid overpressure工况 only)
 * [PUB008] Fault bit3=8: overpressure but no specific cause identified (valid overpressure工况 only)
 * [PUB009] currentCauseMask reset to 0 when NOT runRequest; low 4 bits only; allowed: 0,1,2,4,6,8
 * [PUB010] latchedCauseMask: bitwise OR accumulation while tripLatched=TRUE; cleared on valid reset only
 * [PUB011] fuelPermit = runRequest AND NOT tripLatched; diagnosticActive = currentCauseMask <> 0
 * [PUB012] Output retention: tripLatched holds until valid reset; fuelPermit combinational per PUB011
 * [PUB013] Units: kPa (pressure), t/h (flow), % (valve), dimensionless (bit masks)
 * [PUB014] No hidden timers; all state in VAR; same-scan evaluation per PUB002
 *
 * CONTRACT_RULES [{"kind":"hold_until_reset","output":"tripLatched","set_input":"runRequest","reset_input":"resetBtn"}]
 *)
FUNCTION_BLOCK FB
VAR_INPUT
    runRequest      : BOOL;
    pressure        : REAL;
    pressureValid   : BOOL;
    fuelFlow        : REAL;
    steamFlow       : REAL;
    outletCmd       : INT;
    outletFeedback  : INT;
    resetBtn        : BOOL;
END_VAR
VAR_OUTPUT
    tripLatched     : BOOL;
    fuelPermit      : BOOL;
    currentCauseMask: WORD;
    latchedCauseMask: WORD;
    diagnosticActive: BOOL;
END_VAR
VAR
    prevResetBtn    : BOOL := FALSE;
    prevRunRequest  : BOOL := FALSE;
    stuckCnt        : INT  := 0;
    tempMask        : WORD := 0;
END_VAR

// ---- Rising-edge detection for reset button ----
IF resetBtn AND NOT prevResetBtn THEN
    // Rising edge of resetBtn
    IF NOT runRequest AND pressureValid AND pressure <= 4200.0 THEN
        tripLatched     := FALSE;
        latchedCauseMask := 0;
    END_IF;
END_IF;
prevResetBtn := resetBtn;

// ---- Trip latch activation (PUB002) ----
IF runRequest AND (NOT pressureValid OR pressure >= 4500.0) THEN
    tripLatched := TRUE;
END_IF;

// ---- Fault diagnosis: currentCauseMask (PUB005-PUB009) ----
VAR tempMask : WORD := 0; END_VAR
// bit0: transmitter failure (overrides all other conditions per PUB012)
IF runRequest AND NOT pressureValid THEN
    tempMask := 1; // bit0=1
ELSE
    // bit1 and bit2 only evaluated in valid overpressure工况 (PUB008/PUB009)
    IF runRequest AND pressureValid AND pressure >= 4500.0 THEN
        // Stuck valve counter: 3 consecutive valid scans (PUB006)
        IF outletCmd >= 50 AND outletFeedback <= 10 THEN
            stuckCnt := stuckCnt + 1;
        ELSE
            stuckCnt := 0;
        END_IF;
        IF stuckCnt >= 3 THEN
            tempMask := tempMask OR 2; // bit1=2
        END_IF;
        // Excess combustion: fuelFlow>=4.0 AND steamFlow<=10.0 (PUB007)
        IF fuelFlow >= 4.0 AND steamFlow <= 10.0 THEN
            tempMask := tempMask OR 4; // bit2=4
        END_IF;
        // Unlocated: overpressure but no specific cause (PUB008)
        IF tempMask = 0 THEN
            tempMask := 8; // bit3=8
        END_IF;
    ELSE
        stuckCnt := 0;
    END_IF;
ELSE
    stuckCnt := 0;
END_IF;
currentCauseMask := tempMask;

// ---- Latched cause accumulation (PUB010) ----
IF tripLatched THEN
    latchedCauseMask := latchedCauseMask OR currentCauseMask;
END_IF;

// ---- Fuel permit and diagnostic (PUB011) ----
fuelPermit      := runRequest AND NOT tripLatched;
diagnosticActive := currentCauseMask <> 0;

// ---- Update previous run state for rising-edge tracking ----
prevRunRequest := runRequest;
END_FUNCTION_BLOCK

(* ---- self-hard-06.raw_candidate_03.st ---- *)
(* ENGINEERING_CONTRACT: Steam Header Overpressure Interlock + Fault Diagnosis
 * ================================================================================
 * [PUB001] Function: FB - steam header overpressure interlock with fault footprint
 * [PUB002] Trip activation: runRequest AND (NOT pressureValid OR pressure >= 4500.0) same-scan
 * [PUB003] Reset permission: resetBtn rising-edge AND NOT runRequest AND pressureValid AND pressure <= 4200.0
 * [PUB004] Hysteresis: 300 kPa (4500 trip / 4200 reset gap per PUB003/PUB010)
 * [PUB005] Fault bit0=1: runRequest AND NOT pressureValid (transmitter failure)
 * [PUB006] Fault bit1=2: outletCmd>=50 AND outletFeedback<=10 for 3 consecutive valid overpressure scans
 *            Counter reset on: NOT runRequest, NOT pressureValid, pressure<4500, or condition unsatisfied
 * [PUB007] Fault bit2=4: fuelFlow >= 4.0 AND steamFlow <= 10.0 (valid overpressure工况 only)
 * [PUB008] Fault bit3=8: overpressure but no specific cause identified (valid overpressure工况 only)
 * [PUB009] currentCauseMask reset to 0 when NOT runRequest; low 4 bits only; allowed: 0,1,2,4,6,8
 * [PUB010] latchedCauseMask: bitwise OR accumulation while tripLatched=TRUE; cleared on valid reset only
 * [PUB011] fuelPermit = runRequest AND NOT tripLatched; diagnosticActive = currentCauseMask <> 0
 * [PUB012] Output retention: tripLatched holds until valid reset; fuelPermit combinational per PUB011
 * [PUB013] Units: kPa (pressure), t/h (flow), % (valve), dimensionless (bit masks)
 * [PUB014] No hidden timers; all state in VAR; same-scan evaluation per PUB002
 *
 * CONTRACT_RULES [{"kind":"hold_until_reset","output":"tripLatched","set_input":"runRequest","reset_input":"resetBtn"}]
 *)
FUNCTION_BLOCK FB
VAR_INPUT
    runRequest      : BOOL;
    pressure        : REAL;
    pressureValid   : BOOL;
    fuelFlow        : REAL;
    steamFlow       : REAL;
    outletCmd       : INT;
    outletFeedback  : INT;
    resetBtn        : BOOL;
END_VAR
VAR_OUTPUT
    tripLatched     : BOOL;
    fuelPermit      : BOOL;
    currentCauseMask: WORD;
    latchedCauseMask: WORD;
    diagnosticActive: BOOL;
END_VAR
VAR
    prevResetBtn    : BOOL := FALSE;
    prevRunRequest  : BOOL := FALSE;
    stuckCnt        : INT  := 0;
    tempMask        : WORD := 0;
END_VAR

// ---- Rising-edge detection for reset button ----
IF resetBtn AND NOT prevResetBtn THEN
    IF NOT runRequest AND pressureValid AND pressure <= 4200.0 THEN
        tripLatched      := FALSE;
        latchedCauseMask := 0;
    END_IF;
END_IF;
prevResetBtn := resetBtn;

// ---- Trip latch activation (PUB002) ----
IF runRequest AND (NOT pressureValid OR pressure >= 4500.0) THEN
    tripLatched := TRUE;
END_IF;

// ---- Fault diagnosis: currentCauseMask (PUB005-PUB009) ----
tempMask := 0;
IF runRequest AND NOT pressureValid THEN
    tempMask := 1;
ELSIF runRequest AND pressureValid AND pressure >= 4500.0 THEN
    IF outletCmd >= 50 AND outletFeedback <= 10 THEN
        stuckCnt := stuckCnt + 1;
    ELSE
        stuckCnt := 0;
    END_IF;
    IF stuckCnt >= 3 THEN
        tempMask := tempMask OR 2;
    END_IF;
    IF fuelFlow >= 4.0 AND steamFlow <= 10.0 THEN
        tempMask := tempMask OR 4;
    END_IF;
    IF tempMask = 0 THEN
        tempMask := 8;
    END_IF;
ELSE
    stuckCnt := 0;
END_IF;
currentCauseMask := tempMask;

// ---- Latched cause accumulation (PUB010) ----
IF tripLatched THEN
    latchedCauseMask := latchedCauseMask OR currentCauseMask;
END_IF;

// ---- Fuel permit and diagnostic (PUB011) ----
fuelPermit      := runRequest AND NOT tripLatched;
diagnosticActive := currentCauseMask <> 0;

// ---- Update previous run state for rising-edge tracking ----
prevRunRequest := runRequest;
END_FUNCTION_BLOCK
